(* IEC 61131-3 sources: plc-st-coding-agent/progress/evidence/f14_v3_parallel_20261112/jobs/custom_minimax-m27 (part 2) *)

(* ---- public-hard-06.candidate_01.st ---- *)
FUNCTION_BLOCK ProductionControl
VAR_INPUT
    Mode            : BOOL;
    ForwardButton   : BOOL;
    ReverseButton   : BOOL;
    SensorFeed      : BOOL;
    SensorWash      : BOOL;
    SensorWeight    : BOOL;
    SensorFiring    : BOOL;
    SensorOutput    : BOOL;
    washComplete    : BOOL;
    weightComplete  : BOOL;
    weight          : REAL;
    firingComplete  : BOOL;
END_VAR

VAR_OUTPUT
    MotorForward    : BOOL;
    MotorReverse    : BOOL;
    kick             : BOOL;
    CompletionLight  : BOOL;
    firingTemp       : REAL;
END_VAR

VAR
    State           : INT;
    prevSensorFeed  : BOOL;
    prevSensorWash  : BOOL;
    prevSensorWeight: BOOL;
    prevSensorFiring: BOOL;
    prevSensorOutput: BOOL;
END_VAR

TYPE ProductionState : INT (
    IDLE            := 0,
    MOVING_TO_WASH  := 1,
    AT_WASH         := 2,
    MOVING_TO_WEIGH := 3,
    AT_WEIGH        := 4,
    QUALITY_CHECK   := 5,
    KICKING         := 6,
    CALCULATING_TEMP:= 7,
    MOVING_TO_FIRING:= 8,
    AT_FIRING       := 9,
    MOVING_TO_OUTPUT:= 10,
    AT_OUTPUT       := 11
);
END_TYPE;

// Edge detection helpers
prevSensorFeed  := SensorFeed;
prevSensorWash  := SensorWash;
prevSensorWeight:= SensorWeight;
prevSensorFiring:= SensorFiring;
prevSensorOutput:= SensorOutput;

// Default outputs
MotorForward    := FALSE;
MotorReverse    := FALSE;
kick             := FALSE;
CompletionLight  := FALSE;
firingTemp       := 0.0;

IF Mode = FALSE THEN
    // Manual Mode
    IF ForwardButton AND NOT ReverseButton THEN
        MotorForward := TRUE;
        MotorReverse := FALSE;
    ELSIF ReverseButton AND NOT ForwardButton THEN
        MotorForward := FALSE;
        MotorReverse := TRUE;
    ELSE
        MotorForward := FALSE;
        MotorReverse := FALSE;
    END_IF;
    State := IDLE;
ELSE
    // Automatic Mode
    CASE State OF
        IDLE:
            IF SensorFeed AND NOT prevSensorFeed THEN
                State := MOVING_TO_WASH;
                MotorForward := TRUE;
            END_IF;

        MOVING_TO_WASH:
            IF SensorWash AND NOT prevSensorWash THEN
                State := AT_WASH;
                MotorForward := FALSE;
            END_IF;

        AT_WASH:
            IF washComplete THEN
                State := MOVING_TO_WEIGH;
                MotorForward := TRUE;
            END_IF;

        MOVING_TO_WEIGH:
            IF SensorWeight AND NOT prevSensorWeight THEN
                State := AT_WEIGH;
                MotorForward := FALSE;
            END_IF;

        AT_WEIGH:
            IF weightComplete THEN
                State := QUALITY_CHECK;
            END_IF;

        QUALITY_CHECK:
            IF weight < 100.0 OR weight > 200.0 THEN
                State := KICKING;
            ELSE
                State := CALCULATING_TEMP;
            END_IF;

        KICKING:
            kick := TRUE;
            State := IDLE;

        CALCULATING_TEMP:
            firingTemp := 500.0 + ((weight - 100.0) / 100.0) * 50.0;
            State := MOVING_TO_FIRING;
            MotorForward := TRUE;

        MOVING_TO_FIRING:
            IF SensorFiring AND NOT prevSensorFiring THEN
                State := AT_FIRING;
                MotorForward := FALSE;
            END_IF;

        AT_FIRING:
            IF firingComplete THEN
                State := MOVING_TO_OUTPUT;
                MotorForward := TRUE;
            END_IF;

        MOVING_TO_OUTPUT:
            IF SensorOutput AND NOT prevSensorOutput THEN
                State := AT_OUTPUT;
                MotorForward := FALSE;
            END_IF;

        AT_OUTPUT:
            CompletionLight := SensorOutput;
            IF NOT SensorOutput THEN
                State := IDLE;
                firingTemp := 0.0;
            END_IF;
    END_CASE;
END_IF;
END_FUNCTION_BLOCK

(* ---- public-hard-06.candidate_02.st ---- *)
FUNCTION_BLOCK ProductionControl
VAR_INPUT
    Mode            : BOOL;
    ForwardButton   : BOOL;
    ReverseButton   : BOOL;
    SensorFeed      : BOOL;
    SensorWash      : BOOL;
    SensorWeight    : BOOL;
    SensorFiring    : BOOL;
    SensorOutput    : BOOL;
    washComplete    : BOOL;
    weightComplete  : BOOL;
    weight          : REAL;
    firingComplete  : BOOL;
END_VAR

VAR_OUTPUT
    MotorForward    : BOOL;
    MotorReverse    : BOOL;
    kick             : BOOL;
    CompletionLight  : BOOL;
    firingTemp       : REAL;
END_VAR

VAR
    State           : INT;
    prevSensorFeed  : BOOL;
    prevSensorWash  : BOOL;
    prevSensorWeight: BOOL;
    prevSensorFiring: BOOL;
    prevSensorOutput: BOOL;
    prodState        : INT;
END_VAR

prodState := State;

kick := FALSE;
firingTemp := 0.0;

prevSensorFeed := SensorFeed;
prevSensorWash := SensorWash;
prevSensorWeight := SensorWeight;
prevSensorFiring := SensorFiring;
prevSensorOutput := SensorOutput;

IF Mode = FALSE THEN
    MotorForward := FALSE;
    MotorReverse := FALSE;
    kick := FALSE;
    CompletionLight := FALSE;
    IF ForwardButton AND NOT ReverseButton THEN
        MotorForward := TRUE;
    END_IF;
    IF ReverseButton AND NOT ForwardButton THEN
        MotorReverse := TRUE;
    END_IF;
    State := 0;
ELSE
    CompletionLight := FALSE;
    CASE State OF
        0:
            MotorForward := FALSE;
            MotorReverse := FALSE;
            kick := FALSE;
            IF SensorFeed AND NOT prevSensorFeed THEN
                State := 1;
            END_IF;

        1:
            MotorForward := TRUE;
            MotorReverse := FALSE;
            IF SensorWash AND NOT prevSensorWash THEN
                State := 2;
            END_IF;

        2:
            MotorForward := FALSE;
            MotorReverse := FALSE;
            IF washComplete THEN
                State := 3;
            END_IF;

        3:
            MotorForward := TRUE;
            MotorReverse := FALSE;
            IF SensorWeight AND NOT prevSensorWeight THEN
                State := 4;
            END_IF;

        4:
            MotorForward := FALSE;
            MotorReverse := FALSE;
            IF weightComplete THEN
                State := 5;
            END_IF;

        5:
            MotorForward := FALSE;
            MotorReverse := FALSE;
            IF weight < 100.0 OR weight > 200.0 THEN
                State := 6;
            ELSE
                State := 7;
            END_IF;

        6:
            kick := TRUE;
            MotorForward := FALSE;
            MotorReverse := FALSE;
            State := 0;

        7:
            kick := FALSE;
            firingTemp := 500.0 + ((weight - 100.0) / 100.0) * 50.0;
            State := 8;

        8:
            MotorForward := TRUE;
            MotorReverse := FALSE;
            kick := FALSE;
            IF SensorFiring AND NOT prevSensorFiring THEN
                State := 9;
            END_IF;

        9:
            MotorForward := FALSE;
            MotorReverse := FALSE;
            IF firingComplete THEN
                State := 10;
            END_IF;

        10:
            MotorForward := TRUE;
            MotorReverse := FALSE;
            IF SensorOutput AND NOT prevSensorOutput THEN
                State := 11;
            END_IF;

        11:
            MotorForward := FALSE;
            MotorReverse := FALSE;
            CompletionLight := TRUE;
            IF NOT SensorOutput THEN
                CompletionLight := FALSE;
                firingTemp := 0.0;
                State := 0;
            END_IF;
    END_CASE;
END_IF;
END_FUNCTION_BLOCK

(* ---- public-hard-06.raw_candidate_01.st ---- *)
FUNCTION_BLOCK ProductionControl
VAR_INPUT
    Mode            : BOOL;
    ForwardButton   : BOOL;
    ReverseButton   : BOOL;
    SensorFeed      : BOOL;
    SensorWash      : BOOL;
    SensorWeight    : BOOL;
    SensorFiring    : BOOL;
    SensorOutput    : BOOL;
    washComplete    : BOOL;
    weightComplete  : BOOL;
    weight          : REAL;
    firingComplete  : BOOL;
END_VAR

VAR_OUTPUT
    MotorForward    : BOOL;
    MotorReverse    : BOOL;
    kick             : BOOL;
    CompletionLight  : BOOL;
    firingTemp       : REAL;
END_VAR

VAR
    State           : INT;
    prevSensorFeed  : BOOL;
    prevSensorWash  : BOOL;
    prevSensorWeight: BOOL;
    prevSensorFiring: BOOL;
    prevSensorOutput: BOOL;
END_VAR

TYPE ProductionState : INT (
    IDLE            := 0,
    MOVING_TO_WASH  := 1,
    AT_WASH         := 2,
    MOVING_TO_WEIGH := 3,
    AT_WEIGH        := 4,
    QUALITY_CHECK   := 5,
    KICKING         := 6,
    CALCULATING_TEMP:= 7,
    MOVING_TO_FIRING:= 8,
    AT_FIRING       := 9,
    MOVING_TO_OUTPUT:= 10,
    AT_OUTPUT       := 11
);
END_TYPE

// Edge detection helpers
prevSensorFeed  := SensorFeed;
prevSensorWash  := SensorWash;
prevSensorWeight:= SensorWeight;
prevSensorFiring:= SensorFiring;
prevSensorOutput:= SensorOutput;

// Default outputs
MotorForward    := FALSE;
MotorReverse    := FALSE;
kick             := FALSE;
CompletionLight  := FALSE;
firingTemp       := 0.0;

IF Mode = FALSE THEN
    // Manual Mode
    IF ForwardButton AND NOT ReverseButton THEN
        MotorForward := TRUE;
        MotorReverse := FALSE;
    ELSIF ReverseButton AND NOT ForwardButton THEN
        MotorForward := FALSE;
        MotorReverse := TRUE;
    ELSE
        MotorForward := FALSE;
        MotorReverse := FALSE;
    END_IF;
    State := IDLE;
ELSE
    // Automatic Mode
    CASE State OF
        IDLE:
            IF SensorFeed AND NOT prevSensorFeed THEN
                State := MOVING_TO_WASH;
                MotorForward := TRUE;
            END_IF;

        MOVING_TO_WASH:
            IF SensorWash AND NOT prevSensorWash THEN
                State := AT_WASH;
                MotorForward := FALSE;
            END_IF;

        AT_WASH:
            IF washComplete THEN
                State := MOVING_TO_WEIGH;
                MotorForward := TRUE;
            END_IF;

        MOVING_TO_WEIGH:
            IF SensorWeight AND NOT prevSensorWeight THEN
                State := AT_WEIGH;
                MotorForward := FALSE;
            END_IF;

        AT_WEIGH:
            IF weightComplete THEN
                State := QUALITY_CHECK;
            END_IF;

        QUALITY_CHECK:
            IF weight < 100.0 OR weight > 200.0 THEN
                State := KICKING;
            ELSE
                State := CALCULATING_TEMP;
            END_IF;

        KICKING:
            kick := TRUE;
            State := IDLE;

        CALCULATING_TEMP:
            firingTemp := 500.0 + ((weight - 100.0) / 100.0) * 50.0;
            State := MOVING_TO_FIRING;
            MotorForward := TRUE;

        MOVING_TO_FIRING:
            IF SensorFiring AND NOT prevSensorFiring THEN
                State := AT_FIRING;
                MotorForward := FALSE;
            END_IF;

        AT_FIRING:
            IF firingComplete THEN
                State := MOVING_TO_OUTPUT;
                MotorForward := TRUE;
            END_IF;

        MOVING_TO_OUTPUT:
            IF SensorOutput AND NOT prevSensorOutput THEN
                State := AT_OUTPUT;
                MotorForward := FALSE;
            END_IF;

        AT_OUTPUT:
            CompletionLight := SensorOutput;
            IF NOT SensorOutput THEN
                State := IDLE;
                firingTemp := 0.0;
            END_IF;
    END_CASE;
END_IF;
END_FUNCTION_BLOCK

(* ---- public-hard-06.raw_candidate_02.st ---- *)
FUNCTION_BLOCK ProductionControl
VAR_INPUT
    Mode            : BOOL;
    ForwardButton   : BOOL;
    ReverseButton   : BOOL;
    SensorFeed      : BOOL;
    SensorWash      : BOOL;
    SensorWeight    : BOOL;
    SensorFiring    : BOOL;
    SensorOutput    : BOOL;
    washComplete    : BOOL;
    weightComplete  : BOOL;
    weight          : REAL;
    firingComplete  : BOOL;
END_VAR

VAR_OUTPUT
    MotorForward    : BOOL;
    MotorReverse    : BOOL;
    kick             : BOOL;
    CompletionLight  : BOOL;
    firingTemp       : REAL;
END_VAR

VAR
    State           : INT;
    prevSensorFeed  : BOOL;
    prevSensorWash  : BOOL;
    prevSensorWeight: BOOL;
    prevSensorFiring: BOOL;
    prevSensorOutput: BOOL;
    prodState        : INT;
END_VAR

prodState := State;

kick := FALSE;
firingTemp := 0.0;

prevSensorFeed := SensorFeed;
prevSensorWash := SensorWash;
prevSensorWeight := SensorWeight;
prevSensorFiring := SensorFiring;
prevSensorOutput := SensorOutput;

IF Mode = FALSE THEN
    MotorForward := FALSE;
    MotorReverse := FALSE;
    kick := FALSE;
    CompletionLight := FALSE;
    IF ForwardButton AND NOT ReverseButton THEN
        MotorForward := TRUE;
    END_IF;
    IF ReverseButton AND NOT ForwardButton THEN
        MotorReverse := TRUE;
    END_IF;
    State := 0;
ELSE
    CompletionLight := FALSE;
    CASE State OF
        0:
            MotorForward := FALSE;
            MotorReverse := FALSE;
            kick := FALSE;
            IF SensorFeed AND NOT prevSensorFeed THEN
                State := 1;
            END_IF;

        1:
            MotorForward := TRUE;
            MotorReverse := FALSE;
            IF SensorWash AND NOT prevSensorWash THEN
                State := 2;
            END_IF;

        2:
            MotorForward := FALSE;
            MotorReverse := FALSE;
            IF washComplete THEN
                State := 3;
            END_IF;

        3:
            MotorForward := TRUE;
            MotorReverse := FALSE;
            IF SensorWeight AND NOT prevSensorWeight THEN
                State := 4;
            END_IF;

        4:
            MotorForward := FALSE;
            MotorReverse := FALSE;
            IF weightComplete THEN
                State := 5;
            END_IF;

        5:
            MotorForward := FALSE;
            MotorReverse := FALSE;
            IF weight < 100.0 OR weight > 200.0 THEN
                State := 6;
            ELSE
                State := 7;
            END_IF;

        6:
            kick := TRUE;
            MotorForward := FALSE;
            MotorReverse := FALSE;
            State := 0;

        7:
            kick := FALSE;
            firingTemp := 500.0 + ((weight - 100.0) / 100.0) * 50.0;
            State := 8;

        8:
            MotorForward := TRUE;
            MotorReverse := FALSE;
            kick := FALSE;
            IF SensorFiring AND NOT prevSensorFiring THEN
                State := 9;
            END_IF;

        9:
            MotorForward := FALSE;
            MotorReverse := FALSE;
            IF firingComplete THEN
                State := 10;
            END_IF;

        10:
            MotorForward := TRUE;
            MotorReverse := FALSE;
            IF SensorOutput AND NOT prevSensorOutput THEN
                State := 11;
            END_IF;

        11:
            MotorForward := FALSE;
            MotorReverse := FALSE;
            CompletionLight := TRUE;
            IF NOT SensorOutput THEN
                CompletionLight := FALSE;
                firingTemp := 0.0;
                State := 0;
            END_IF;
    END_CASE;
END_IF;
END_FUNCTION_BLOCK

(* ---- public-medium-01.candidate_01.st ---- *)
FUNCTION_BLOCK FB_MultiPumpControl
VAR_INPUT
    mode  : BOOL;    // FALSE: Manual, TRUE: Automatic
    start : BOOL;    // Start button
    stop  : BOOL;    // Stop button
END_VAR

VAR_IN_OUT
    pumpGroup : ARRAY[1..5] OF ST_Pump;
END_VAR

VAR
    lastStart : BOOL := FALSE;
    lastStop  : BOOL := FALSE;
    edgeStart : BOOL;
    edgeStop  : BOOL;
    i         : INT;
    j         : INT;
    tempPri   : INT;
    tempSel   : BOOL;
    tempCmd   : BOOL;
    sorted    : ARRAY[1..5] OF ST_Pump;
END_VAR

// Edge detection for rising edges
edgeStart := start AND NOT lastStart;
edgeStop  := stop  AND NOT lastStop;
lastStart := start;
lastStop  := stop;

// Stop all pumps when stop button is pressed
IF edgeStop THEN
    FOR i := 1 TO 5 DO
        pumpGroup[i].RunComd := FALSE;
    END_FOR;
END_IF;

// Start selected pumps when start button is pressed
IF edgeStart THEN
    IF mode = FALSE THEN
        // Manual mode: run pumps where selection = TRUE
        FOR i := 1 TO 5 DO
            pumpGroup[i].RunComd := pumpGroup[i].selection;
        END_FOR;
    ELSE
        // Automatic mode: three pumps in use, two on standby
        // Sort pumps by priority (descending) using bubble sort
        sorted := pumpGroup;
        FOR i := 1 TO 4 DO
            FOR j := 1 TO 5 - i DO
                IF sorted[j].priority < sorted[j + 1].priority THEN
                    tempPri := sorted[j].priority;
                    tempSel := sorted[j].selection;
                    tempCmd := sorted[j].RunComd;
                    sorted[j].priority   := sorted[j + 1].priority;
                    sorted[j].selection  := sorted[j + 1].selection;
                    sorted[j].RunComd    := sorted[j + 1].RunComd;
                    sorted[j + 1].priority := tempPri;
                    sorted[j + 1].selection := tempSel;
                    sorted[j + 1].RunComd   := tempCmd;
                END_IF;
            END_FOR;
        END_FOR;
        // Top 3 highest priority pumps run
        sorted[1].RunComd := TRUE;
        sorted[2].RunComd := TRUE;
        sorted[3].RunComd := TRUE;
        sorted[4].RunComd := FALSE;
        sorted[5].RunComd := FALSE;
        // Copy RunComd back to original array (preserving original order)
        FOR i := 1 TO 5 DO
            pumpGroup[i].RunComd := sorted[i].RunComd;
        END_FOR;
    END_IF;
END_IF;

END_FUNCTION_BLOCK

(* ---- public-medium-01.candidate_02.st ---- *)
TYPE ST_Pump : STRUCT
    priority : INT;
    selection : BOOL;
    runCmd   : BOOL;
END_STRUCT;
END_TYPE;

FUNCTION_BLOCK FB_MultiPumpControl
VAR_INPUT
    mode  : BOOL;
    start : BOOL;
    stop  : BOOL;
END_VAR

VAR_IN_OUT
    pumpGroup : ARRAY[1..5] OF ST_Pump;
END_VAR

VAR
    lastStart : BOOL := FALSE;
    lastStop  : BOOL := FALSE;
    edgeStart : BOOL;
    edgeStop  : BOOL;
    i         : INT;
    j         : INT;
    tempPump  : ST_Pump;
    pumpSorted : ARRAY[1..5] OF ST_Pump;
END_VAR

edgeStart := start AND NOT lastStart;
edgeStop  := stop  AND NOT lastStop;
lastStart := start;
lastStop  := stop;

IF edgeStop THEN
    FOR i := 1 TO 5 DO
        pumpGroup[i].runCmd := FALSE;
    END_FOR;
END_IF;

IF edgeStart THEN
    IF mode = FALSE THEN
        FOR i := 1 TO 5 DO
            pumpGroup[i].runCmd := pumpGroup[i].selection;
        END_FOR;
    ELSE
        pumpSorted := pumpGroup;
        FOR i := 1 TO 4 DO
            FOR j := 1 TO 5 - i DO
                IF pumpSorted[j].priority < pumpSorted[j + 1].priority THEN
                    tempPump := pumpSorted[j];
                    pumpSorted[j] := pumpSorted[j + 1];
                    pumpSorted[j + 1] := tempPump;
                END_IF;
            END_FOR;
        END_FOR;
        pumpSorted[1].runCmd := TRUE;
        pumpSorted[2].runCmd := TRUE;
        pumpSorted[3].runCmd := TRUE;
        pumpSorted[4].runCmd := FALSE;
        pumpSorted[5].runCmd := FALSE;
        pumpGroup := pumpSorted;
    END_IF;
END_IF;

END_FUNCTION_BLOCK

(* ---- public-medium-01.raw_candidate_01.st ---- *)
FUNCTION_BLOCK FB_MultiPumpControl
VAR_INPUT
    mode  : BOOL;    // FALSE: Manual, TRUE: Automatic
    start : BOOL;    // Start button
    stop  : BOOL;    // Stop button
END_VAR

VAR_IN_OUT
    pumpGroup : ARRAY[1..5] OF ST_Pump;
END_VAR

VAR
    lastStart : BOOL := FALSE;
    lastStop  : BOOL := FALSE;
    edgeStart : BOOL;
    edgeStop  : BOOL;
    i         : INT;
    j         : INT;
    tempPri   : INT;
    tempSel   : BOOL;
    tempCmd   : BOOL;
    sorted    : ARRAY[1..5] OF ST_Pump;
END_VAR

// Edge detection for rising edges
edgeStart := start AND NOT lastStart;
edgeStop  := stop  AND NOT lastStop;
lastStart := start;
lastStop  := stop;

// Stop all pumps when stop button is pressed
IF edgeStop THEN
    FOR i := 1 TO 5 DO
        pumpGroup[i].RunComd := FALSE;
    END_FOR;
END_IF

// Start selected pumps when start button is pressed
IF edgeStart THEN
    IF mode = FALSE THEN
        // Manual mode: run pumps where selection = TRUE
        FOR i := 1 TO 5 DO
            pumpGroup[i].RunComd := pumpGroup[i].selection;
        END_FOR;
    ELSE
        // Automatic mode: three pumps in use, two on standby
        // Sort pumps by priority (descending) using bubble sort
        sorted := pumpGroup;
        FOR i := 1 TO 4 DO
            FOR j := 1 TO 5 - i DO
                IF sorted[j].priority < sorted[j + 1].priority THEN
                    tempPri := sorted[j].priority;
                    tempSel := sorted[j].selection;
                    tempCmd := sorted[j].RunComd;
                    sorted[j].priority   := sorted[j + 1].priority;
                    sorted[j].selection  := sorted[j + 1].selection;
                    sorted[j].RunComd    := sorted[j + 1].RunComd;
                    sorted[j + 1].priority := tempPri;
                    sorted[j + 1].selection := tempSel;
                    sorted[j + 1].RunComd   := tempCmd;
                END_IF
            END_FOR
        END_FOR
        // Top 3 highest priority pumps run
        sorted[1].RunComd := TRUE;
        sorted[2].RunComd := TRUE;
        sorted[3].RunComd := TRUE;
        sorted[4].RunComd := FALSE;
        sorted[5].RunComd := FALSE;
        // Copy RunComd back to original array (preserving original order)
        FOR i := 1 TO 5 DO
            pumpGroup[i].RunComd := sorted[i].RunComd;
        END_FOR;
    END_IF
END_IF

END_FUNCTION_BLOCK

(* ---- public-medium-01.raw_candidate_02.st ---- *)
TYPE ST_Pump : STRUCT
    priority : INT;
    selection : BOOL;
    runCmd   : BOOL;
END_STRUCT
END_TYPE

FUNCTION_BLOCK FB_MultiPumpControl
VAR_INPUT
    mode  : BOOL;
    start : BOOL;
    stop  : BOOL;
END_VAR

VAR_IN_OUT
    pumpGroup : ARRAY[1..5] OF ST_Pump;
END_VAR

VAR
    lastStart : BOOL := FALSE;
    lastStop  : BOOL := FALSE;
    edgeStart : BOOL;
    edgeStop  : BOOL;
    i         : INT;
    j         : INT;
    tempPump  : ST_Pump;
    pumpSorted : ARRAY[1..5] OF ST_Pump;
END_VAR

edgeStart := start AND NOT lastStart;
edgeStop  := stop  AND NOT lastStop;
lastStart := start;
lastStop  := stop;

IF edgeStop THEN
    FOR i := 1 TO 5 DO
        pumpGroup[i].runCmd := FALSE;
    END_FOR;
END_IF;

IF edgeStart THEN
    IF mode = FALSE THEN
        FOR i := 1 TO 5 DO
            pumpGroup[i].runCmd := pumpGroup[i].selection;
        END_FOR;
    ELSE
        pumpSorted := pumpGroup;
        FOR i := 1 TO 4 DO
            FOR j := 1 TO 5 - i DO
                IF pumpSorted[j].priority < pumpSorted[j + 1].priority THEN
                    tempPump := pumpSorted[j];
                    pumpSorted[j] := pumpSorted[j + 1];
                    pumpSorted[j + 1] := tempPump;
                END_IF;
            END_FOR;
        END_FOR;
        pumpSorted[1].runCmd := TRUE;
        pumpSorted[2].runCmd := TRUE;
        pumpSorted[3].runCmd := TRUE;
        pumpSorted[4].runCmd := FALSE;
        pumpSorted[5].runCmd := FALSE;
        pumpGroup := pumpSorted;
    END_IF;
END_IF;

END_FUNCTION_BLOCK

(* ---- public-medium-02.candidate_01.st ---- *)
FUNCTION_BLOCK FB_AnalogBatchProcessing
VAR_INPUT
    count : DINT;
END_VAR

VAR_IN_OUT
    analogValues : ARRAY[*] OF INT;
    channels : ARRAY[*] OF ST_AnalogChannel;
END_VAR

VAR
    i : DINT;
    idx : DINT;
    rawValue : INT;
    rawMin : INT;
    rawMax : INT;
    loLIM : REAL;
    hiLIM : REAL;
END_VAR

loLIM := 0.0;
hiLIM := 0.0;

FOR i := 0 TO count - 1 DO
    idx := LOWER_BOUND(analogValues, 1) + i;
    rawValue := analogValues[idx];

    channels[idx].retVal := 16#0000;

    IF channels[idx].enable THEN
        loLIM := channels[idx].loLIM;
        hiLIM := channels[idx].hiLIM;

        CASE channels[idx].measuringMode OF
            0: // Non-temperature linear scaling
                IF hiLIM > loLIM THEN
                    IF channels[idx].bipolar THEN
                        rawMin := -27648;
                        rawMax := 27648;
                    ELSE
                        rawMin := 0;
                        rawMax := 27648;
                    END_IF;

                    channels[idx].outputValue := TO_REAL(rawValue - rawMin) / TO_REAL(rawMax - rawMin) * (hiLIM - loLIM) + loLIM;
                ELSE
                    channels[idx].retVal := 16#8002;
                END_IF;

            1: // Standard temperature: outputValue = raw / 10
                channels[idx].outputValue := TO_REAL(rawValue) / 10.0;

            2: // Climatic temperature: outputValue = raw / 100
                channels[idx].outputValue := TO_REAL(rawValue) / 100.0;

            ELSE
                channels[idx].retVal := 16#8001;
        END_CASE;
    END_IF;
END_FOR;
END_FUNCTION_BLOCK

(* ---- public-medium-02.candidate_02.st ---- *)
TYPE ST_AnalogChannel :
STRUCT
    enable : BOOL;
    hiLIM : REAL;
    loLIM : REAL;
    bipolar : BOOL;
    measuringMode : INT;
    retVal : WORD;
    outputValue : REAL;
END_STRUCT;
END_TYPE;

FUNCTION_BLOCK FB_AnalogBatchProcessing
VAR_INPUT
    count : DINT;
END_VAR

VAR_IN_OUT
    analogValues : ARRAY[*] OF INT;
    channels : ARRAY[*] OF ST_AnalogChannel;
END_VAR

VAR
    i : DINT;
    idx : DINT;
    rawValue : INT;
    rawMin : INT;
    rawMax : INT;
    chLoLIM : REAL;
    chHiLIM : REAL;
    ch : REFERENCE TO ST_AnalogChannel;
END_VAR

FOR i := 0 TO count - 1 DO
    idx := LOWER_BOUND(analogValues, 1) + i;
    rawValue := analogValues[idx];
    ch REF= channels[idx];
    ch.retVal := 16#0000;

    IF ch.enable THEN
        chLoLIM := ch.loLIM;
        chHiLIM := ch.hiLIM;

        CASE ch.measuringMode OF
            0:
                IF chHiLIM > chLoLIM THEN
                    IF ch.bipolar THEN
                        rawMin := -27648;
                        rawMax := 27648;
                    ELSE
                        rawMin := 0;
                        rawMax := 27648;
                    END_IF;
                    ch.outputValue := INT_TO_REAL(rawValue - rawMin) / INT_TO_REAL(rawMax - rawMin) * (chHiLIM - chLoLIM) + chLoLIM;
                ELSE
                    ch.retVal := 16#8002;
                END_IF;

            1:
                ch.outputValue := INT_TO_REAL(rawValue) / 10.0;

            2:
                ch.outputValue := INT_TO_REAL(rawValue) / 100.0;

            ELSE
                ch.retVal := 16#8001;
        END_CASE;
    END_IF;
END_FOR;
END_FUNCTION_BLOCK

(* ---- public-medium-02.raw_candidate_01.st ---- *)
FUNCTION_BLOCK FB_AnalogBatchProcessing
VAR_INPUT
    count : DINT;
END_VAR

VAR_IN_OUT
    analogValues : ARRAY[*] OF INT;
    channels : ARRAY[*] OF ST_AnalogChannel;
END_VAR

VAR
    i : DINT;
    idx : DINT;
    rawValue : INT;
    rawMin : INT;
    rawMax : INT;
    loLIM : REAL;
    hiLIM : REAL;
END_VAR

loLIM := 0.0;
hiLIM := 0.0;

FOR i := 0 TO count - 1 DO
    idx := LOWER_BOUND(analogValues, 1) + i;
    rawValue := analogValues[idx];

    channels[idx].retVal := 16#0000;

    IF channels[idx].enable THEN
        loLIM := channels[idx].loLIM;
        hiLIM := channels[idx].hiLIM;

        CASE channels[idx].measuringMode OF
            0: // Non-temperature linear scaling
                IF hiLIM > loLIM THEN
                    IF channels[idx].bipolar THEN
                        rawMin := -27648;
                        rawMax := 27648;
                    ELSE
                        rawMin := 0;
                        rawMax := 27648;
                    END_IF;

                    channels[idx].outputValue := TO_REAL(rawValue - rawMin) / TO_REAL(rawMax - rawMin) * (hiLIM - loLIM) + loLIM;
                ELSE
                    channels[idx].retVal := 16#8002;
                END_IF;

            1: // Standard temperature: outputValue = raw / 10
                channels[idx].outputValue := TO_REAL(rawValue) / 10.0;

            2: // Climatic temperature: outputValue = raw / 100
                channels[idx].outputValue := TO_REAL(rawValue) / 100.0;

            ELSE
                channels[idx].retVal := 16#8001;
        END_CASE;
    END_IF;
END_FOR;
END_FUNCTION_BLOCK

(* ---- public-medium-02.raw_candidate_02.st ---- *)
TYPE ST_AnalogChannel :
STRUCT
    enable : BOOL;
    hiLIM : REAL;
    loLIM : REAL;
    bipolar : BOOL;
    measuringMode : INT;
    retVal : WORD;
    outputValue : REAL;
END_STRUCT
END_TYPE

FUNCTION_BLOCK FB_AnalogBatchProcessing
VAR_INPUT
    count : DINT;
END_VAR

VAR_IN_OUT
    analogValues : ARRAY[*] OF INT;
    channels : ARRAY[*] OF ST_AnalogChannel;
END_VAR

VAR
    i : DINT;
    idx : DINT;
    rawValue : INT;
    rawMin : INT;
    rawMax : INT;
    chLoLIM : REAL;
    chHiLIM : REAL;
    ch : REFERENCE TO ST_AnalogChannel;
END_VAR

FOR i := 0 TO count - 1 DO
    idx := LOWER_BOUND(analogValues, 1) + i;
    rawValue := analogValues[idx];
    ch REF= channels[idx];
    ch.retVal := 16#0000;

    IF ch.enable THEN
        chLoLIM := ch.loLIM;
        chHiLIM := ch.hiLIM;

        CASE ch.measuringMode OF
            0:
                IF chHiLIM > chLoLIM THEN
                    IF ch.bipolar THEN
                        rawMin := -27648;
                        rawMax := 27648;
                    ELSE
                        rawMin := 0;
                        rawMax := 27648;
                    END_IF;
                    ch.outputValue := INT_TO_REAL(rawValue - rawMin) / INT_TO_REAL(rawMax - rawMin) * (chHiLIM - chLoLIM) + chLoLIM;
                ELSE
                    ch.retVal := 16#8002;
                END_IF;

            1:
                ch.outputValue := INT_TO_REAL(rawValue) / 10.0;

            2:
                ch.outputValue := INT_TO_REAL(rawValue) / 100.0;

            ELSE
                ch.retVal := 16#8001;
        END_CASE;
    END_IF;
END_FOR;
END_FUNCTION_BLOCK

(* ---- public-medium-03.candidate_01.st ---- *)
FUNCTION_BLOCK FB_MovingAverage
VAR_INPUT
    cyclicExecution : BOOL;
    trigger : BOOL;
    value : LREAL;
    windowSize : INT;
    reset : BOOL;
END_VAR

VAR_OUTPUT
    average : LREAL;
    windowSizeReached : BOOL;
    error : BOOL;
    status : WORD;
END_VAR

VAR
    dataBuffer : ARRAY[1..100] OF LREAL;
    sum : LREAL;
    count : INT;
    writeIndex : INT;
    lastTrigger : BOOL;
    lastReset : BOOL;
    initValid : BOOL;
END_VAR

// Reset handling
IF reset AND NOT lastReset THEN
    sum := 0.0;
    count := 0;
    writeIndex := 0;
    average := 0.0;
    windowSizeReached := FALSE;
    error := FALSE;
    status := 16#0000;
    initValid := FALSE;
END_IF;
lastReset := reset;

// Validate window size on first execution or when reset was just released
IF NOT initValid THEN
    IF windowSize < 1 OR windowSize > 100 THEN
        error := TRUE;
        status := 16#8200;
        RETURN;
    ELSE
        error := FALSE;
        status := 16#0000;
        initValid := TRUE;
    END_IF;
END_IF;

// Check for cyclic execution mode
IF cyclicExecution THEN
    // Validate window size on each cycle
    IF windowSize < 1 OR windowSize > 100 THEN
        error := TRUE;
        status := 16#8200;
        RETURN;
    ELSE
        error := FALSE;
        status := 16#0000;
    END_IF;

    // Process new value
    IF count >= windowSize THEN
        sum := sum - dataBuffer[writeIndex + 1];
    ELSE
        count := count + 1;
    END_IF;

    writeIndex := (writeIndex MOD windowSize) + 1;
    dataBuffer[writeIndex] := value;
    sum := sum + value;

    IF count >= windowSize THEN
        windowSizeReached := TRUE;
    ELSE
        windowSizeReached := FALSE;
    END_IF;

    average := sum / INT_TO_LREAL(count);
    lastTrigger := FALSE;
    RETURN;
END_IF;

// Check for rising edge on trigger
IF trigger AND NOT lastTrigger THEN
    // Validate window size
    IF windowSize < 1 OR windowSize > 100 THEN
        error := TRUE;
        status := 16#8200;
        lastTrigger := trigger;
        RETURN;
    ELSE
        error := FALSE;
        status := 16#0000;
    END_IF;

    // Process new value
    IF count >= windowSize THEN
        sum := sum - dataBuffer[writeIndex + 1];
    ELSE
        count := count + 1;
    END_IF;

    writeIndex := (writeIndex MOD windowSize) + 1;
    dataBuffer[writeIndex] := value;
    sum := sum + value;

    IF count >= windowSize THEN
        windowSizeReached := TRUE;
    ELSE
        windowSizeReached := FALSE;
    END_IF;

    average := sum / INT_TO_LREAL(count);
END_IF;

lastTrigger := trigger;
END_FUNCTION_BLOCK

(* ---- public-medium-03.candidate_02.st ---- *)
FUNCTION_BLOCK FB_MovingAverage
VAR_INPUT
    cyclicExecution : BOOL;
    trigger : BOOL;
    value : LREAL;
    windowSize : INT;
    reset : BOOL;
END_VAR

VAR_OUTPUT
    average : LREAL;
    windowSizeReached : BOOL;
    error : BOOL;
    status : WORD;
END_VAR

VAR
    dataBuffer : ARRAY[1..100] OF LREAL;
    sum : LREAL;
    count : INT;
    writeIndex : INT;
    lastTrigger : BOOL;
    lastReset : BOOL;
    initValid : BOOL;
END_VAR

IF reset AND NOT lastReset THEN
    sum := 0.0;
    count := 0;
    writeIndex := 0;
    average := 0.0;
    windowSizeReached := FALSE;
    error := FALSE;
    status := 16#0000;
    initValid := FALSE;
END_IF;
lastReset := reset;

IF NOT initValid THEN
    IF windowSize < 1 OR windowSize > 100 THEN
        error := TRUE;
        status := 16#8200;
        RETURN;
    ELSE
        error := FALSE;
        status := 16#0000;
        initValid := TRUE;
    END_IF;
END_IF;

IF cyclicExecution THEN
    IF windowSize < 1 OR windowSize > 100 THEN
        error := TRUE;
        status := 16#8200;
        RETURN;
    ELSE
        error := FALSE;
        status := 16#0000;
    END_IF;

    IF count >= windowSize THEN
        sum := sum - dataBuffer[((writeIndex) MOD windowSize) + 1];
    ELSE
        count := count + 1;
    END_IF;

    writeIndex := writeIndex + 1;
    IF writeIndex > windowSize THEN
        writeIndex := 1;
    END_IF;

    dataBuffer[writeIndex] := value;
    sum := sum + value;

    IF count >= windowSize THEN
        windowSizeReached := TRUE;
        average := sum / INT_TO_LREAL(windowSize);
    ELSE
        windowSizeReached := FALSE;
        average := sum / INT_TO_LREAL(count);
    END_IF;
    lastTrigger := FALSE;
    RETURN;
END_IF;

IF trigger AND NOT lastTrigger THEN
    IF windowSize < 1 OR windowSize > 100 THEN
        error := TRUE;
        status := 16#8200;
        lastTrigger := trigger;
        RETURN;
    ELSE
        error := FALSE;
        status := 16#0000;
    END_IF;

    IF count >= windowSize THEN
        sum := sum - dataBuffer[((writeIndex) MOD windowSize) + 1];
    ELSE
        count := count + 1;
    END_IF;

    writeIndex := writeIndex + 1;
    IF writeIndex > windowSize THEN
        writeIndex := 1;
    END_IF;

    dataBuffer[writeIndex] := value;
    sum := sum + value;

    IF count >= windowSize THEN
        windowSizeReached := TRUE;
        average := sum / INT_TO_LREAL(windowSize);
    ELSE
        windowSizeReached := FALSE;
        average := sum / INT_TO_LREAL(count);
    END_IF;
END_IF;

lastTrigger := trigger;
END_FUNCTION_BLOCK

(* ---- public-medium-03.raw_candidate_01.st ---- *)
FUNCTION_BLOCK FB_MovingAverage
VAR_INPUT
    cyclicExecution : BOOL;
    trigger : BOOL;
    value : LREAL;
    windowSize : INT;
    reset : BOOL;
END_VAR

VAR_OUTPUT
    average : LREAL;
    windowSizeReached : BOOL;
    error : BOOL;
    status : WORD;
END_VAR

VAR
    dataBuffer : ARRAY[1..100] OF LREAL;
    sum : LREAL;
    count : INT;
    writeIndex : INT;
    lastTrigger : BOOL;
    lastReset : BOOL;
    initValid : BOOL;
END_VAR

// Reset handling
IF reset AND NOT lastReset THEN
    sum := 0.0;
    count := 0;
    writeIndex := 0;
    average := 0.0;
    windowSizeReached := FALSE;
    error := FALSE;
    status := 16#0000;
    initValid := FALSE;
END_IF;
lastReset := reset;

// Validate window size on first execution or when reset was just released
IF NOT initValid THEN
    IF windowSize < 1 OR windowSize > 100 THEN
        error := TRUE;
        status := 16#8200;
        RETURN;
    ELSE
        error := FALSE;
        status := 16#0000;
        initValid := TRUE;
    END_IF;
END_IF;

// Check for cyclic execution mode
IF cyclicExecution THEN
    // Validate window size on each cycle
    IF windowSize < 1 OR windowSize > 100 THEN
        error := TRUE;
        status := 16#8200;
        RETURN;
    ELSE
        error := FALSE;
        status := 16#0000;
    END_IF;

    // Process new value
    IF count >= windowSize THEN
        sum := sum - dataBuffer[writeIndex + 1];
    ELSE
        count := count + 1;
    END_IF;

    writeIndex := (writeIndex MOD windowSize) + 1;
    dataBuffer[writeIndex] := value;
    sum := sum + value;

    IF count >= windowSize THEN
        windowSizeReached := TRUE;
    ELSE
        windowSizeReached := FALSE;
    END_IF;

    average := sum / INT_TO_LREAL(count);
    lastTrigger := FALSE;
    RETURN;
END_IF;

// Check for rising edge on trigger
IF trigger AND NOT lastTrigger THEN
    // Validate window size
    IF windowSize < 1 OR windowSize > 100 THEN
        error := TRUE;
        status := 16#8200;
        lastTrigger := trigger;
        RETURN;
    ELSE
        error := FALSE;
        status := 16#0000;
    END_IF;

    // Process new value
    IF count >= windowSize THEN
        sum := sum - dataBuffer[writeIndex + 1];
    ELSE
        count := count + 1;
    END_IF;

    writeIndex := (writeIndex MOD windowSize) + 1;
    dataBuffer[writeIndex] := value;
    sum := sum + value;

    IF count >= windowSize THEN
        windowSizeReached := TRUE;
    ELSE
        windowSizeReached := FALSE;
    END_IF;

    average := sum / INT_TO_LREAL(count);
END_IF;

lastTrigger := trigger;
END_FUNCTION_BLOCK

(* ---- public-medium-03.raw_candidate_02.st ---- *)
FUNCTION_BLOCK FB_MovingAverage
VAR_INPUT
    cyclicExecution : BOOL;
    trigger : BOOL;
    value : LREAL;
    windowSize : INT;
    reset : BOOL;
END_VAR

VAR_OUTPUT
    average : LREAL;
    windowSizeReached : BOOL;
    error : BOOL;
    status : WORD;
END_VAR

VAR
    dataBuffer : ARRAY[1..100] OF LREAL;
    sum : LREAL;
    count : INT;
    writeIndex : INT;
    lastTrigger : BOOL;
    lastReset : BOOL;
    initValid : BOOL;
END_VAR

IF reset AND NOT lastReset THEN
    sum := 0.0;
    count := 0;
    writeIndex := 0;
    average := 0.0;
    windowSizeReached := FALSE;
    error := FALSE;
    status := 16#0000;
    initValid := FALSE;
END_IF;
lastReset := reset;

IF NOT initValid THEN
    IF windowSize < 1 OR windowSize > 100 THEN
        error := TRUE;
        status := 16#8200;
        RETURN;
    ELSE
        error := FALSE;
        status := 16#0000;
        initValid := TRUE;
    END_IF;
END_IF;

IF cyclicExecution THEN
    IF windowSize < 1 OR windowSize > 100 THEN
        error := TRUE;
        status := 16#8200;
        RETURN;
    ELSE
        error := FALSE;
        status := 16#0000;
    END_IF;

    IF count >= windowSize THEN
        sum := sum - dataBuffer[((writeIndex) MOD windowSize) + 1];
    ELSE
        count := count + 1;
    END_IF;

    writeIndex := writeIndex + 1;
    IF writeIndex > windowSize THEN
        writeIndex := 1;
    END_IF;

    dataBuffer[writeIndex] := value;
    sum := sum + value;

    IF count >= windowSize THEN
        windowSizeReached := TRUE;
        average := sum / INT_TO_LREAL(windowSize);
    ELSE
        windowSizeReached := FALSE;
        average := sum / INT_TO_LREAL(count);
    END_IF;
    lastTrigger := FALSE;
    RETURN;
END_IF;

IF trigger AND NOT lastTrigger THEN
    IF windowSize < 1 OR windowSize > 100 THEN
        error := TRUE;
        status := 16#8200;
        lastTrigger := trigger;
        RETURN;
    ELSE
        error := FALSE;
        status := 16#0000;
    END_IF;

    IF count >= windowSize THEN
        sum := sum - dataBuffer[((writeIndex) MOD windowSize) + 1];
    ELSE
        count := count + 1;
    END_IF;

    writeIndex := writeIndex + 1;
    IF writeIndex > windowSize THEN
        writeIndex := 1;
    END_IF;

    dataBuffer[writeIndex] := value;
    sum := sum + value;

    IF count >= windowSize THEN
        windowSizeReached := TRUE;
        average := sum / INT_TO_LREAL(windowSize);
    ELSE
        windowSizeReached := FALSE;
        average := sum / INT_TO_LREAL(count);
    END_IF;
END_IF;

lastTrigger := trigger;
END_FUNCTION_BLOCK

(* ---- public-medium-04.candidate_01.st ---- *)
FUNCTION_BLOCK FB_TemperatureControl
VAR_INPUT
    TemperatureSensorInput : REAL;
    SetTemperature : REAL;
END_VAR
VAR_OUTPUT
    CurrentTemperature : REAL;
    SetTempDisplay : REAL;
    HeaterStatus : BOOL;
    OverheatProtection : BOOL;
    HeaterOutput : BOOL;
END_VAR
VAR
    OverheatTimer : TON;
    LockoutTimer : TON;
    OverheatTriggered : BOOL := FALSE;
    LockoutActive : BOOL := FALSE;
END_VAR

(* Constants *)
OverheatTimer.PT := T#5S;
LockoutTimer.PT := T#3S;

(* Sensor fault check: temperature out of valid range *)
IF TemperatureSensorInput < 0.0 OR TemperatureSensorInput > 100.0 THEN
    HeaterOutput := FALSE;
    OverheatTimer(IN := FALSE);
    LockoutTimer(IN := FALSE);
    LockoutActive := FALSE;
    OverheatTriggered := FALSE;
ELSE
    (* Normal temperature control *)

    (* Start overheat timer when heater is commanded ON *)
    OverheatTimer(IN := TRUE);

    (* Check if overheat timer exceeded 5s → trigger protection *)
    IF OverheatTimer.Q AND NOT OverheatTriggered THEN
        OverheatTriggered := TRUE;
        LockoutActive := TRUE;
        LockoutTimer(IN := TRUE);
    END_IF;

    (* If protection triggered, force heater OFF and wait lockout *)
    IF OverheatTriggered THEN
        HeaterOutput := FALSE;

        (* After lockout expires, clear protection *)
        IF LockoutTimer.Q THEN
            LockoutActive := FALSE;
            OverheatTriggered := FALSE;
            LockoutTimer(IN := FALSE);
            OverheatTimer(IN := FALSE);
        END_IF;
    ELSE
        (* Normal operation: compare temperature vs setpoint *)
        IF TemperatureSensorInput < SetTemperature THEN
            HeaterOutput := TRUE;
        ELSE
            HeaterOutput := FALSE;
        END_IF;
    END_IF;

    (* Reset overheat timer when heater is OFF (but not in protection) *)
    IF NOT HeaterOutput AND NOT OverheatTriggered THEN
        OverheatTimer(IN := FALSE);
    END_IF;
END_IF;

(* Update display outputs *)
CurrentTemperature := TemperatureSensorInput;
SetTempDisplay := SetTemperature;
HeaterStatus := HeaterOutput;
OverheatProtection := OverheatTriggered;

END_FUNCTION_BLOCK

(* ---- public-medium-04.candidate_02.st ---- *)
FUNCTION_BLOCK FB_TemperatureControl
VAR_INPUT
    TemperatureSensorInput : REAL;
    SetTemperature : REAL;
END_VAR
VAR_OUTPUT
    CurrentTemperature : REAL;
    SetTempDisplay : REAL;
    HeaterStatus : BOOL;
    OverheatProtection : BOOL;
    HeaterOutput : BOOL;
END_VAR
VAR
    OverheatTimer : TON;
    LockoutTimer : TON;
    OverheatTriggered : BOOL := FALSE;
END_VAR

OverheatTimer.PT := T#5S;
LockoutTimer.PT := T#3S;

(* Sensor fault check: temperature out of valid range *)
IF TemperatureSensorInput < 0.0 OR TemperatureSensorInput > 100.0 THEN
    HeaterOutput := FALSE;
    OverheatTimer(IN := FALSE);
    LockoutTimer(IN := FALSE);
    OverheatTimer(IN := FALSE, PT := T#5S);
    OverheatTriggered := FALSE;
ELSE
    (* Normal temperature control *)
    IF NOT OverheatTriggered THEN
        (* Normal heating decision *)
        IF TemperatureSensorInput < SetTemperature THEN
            HeaterOutput := TRUE;
        ELSE
            HeaterOutput := FALSE;
        END_IF;
    ELSE
        (* Overheat protection active - heater forced off *)
        HeaterOutput := FALSE;
    END_IF;

    (* Overheat timer: accumulate time only when heater is ON and not in protection *)
    IF NOT OverheatTriggered AND HeaterOutput THEN
        OverheatTimer(IN := TRUE);
    ELSE
        OverheatTimer(IN := FALSE);
    END_IF;

    (* Check overheat threshold *)
    IF OverheatTimer.Q AND NOT OverheatTriggered THEN
        OverheatTriggered := TRUE;
    END_IF;

    (* Lockout timer management *)
    IF OverheatTriggered THEN
        LockoutTimer(IN := TRUE);
        IF LockoutTimer.Q THEN
            OverheatTriggered := FALSE;
            LockoutTimer(IN := FALSE);
            OverheatTimer(IN := FALSE, PT := T#5S);
        END_IF;
    ELSE
        LockoutTimer(IN := FALSE);
    END_IF;
END_IF;

(* Update display outputs *)
CurrentTemperature := TemperatureSensorInput;
SetTempDisplay := SetTemperature;
HeaterStatus := HeaterOutput;
OverheatProtection := OverheatTriggered;

END_FUNCTION_BLOCK

(* ---- public-medium-04.raw_candidate_01.st ---- *)
FUNCTION_BLOCK FB_TemperatureControl
VAR_INPUT
    TemperatureSensorInput : REAL;
    SetTemperature : REAL;
END_VAR
VAR_OUTPUT
    CurrentTemperature : REAL;
    SetTempDisplay : REAL;
    HeaterStatus : BOOL;
    OverheatProtection : BOOL;
    HeaterOutput : BOOL;
END_VAR
VAR
    OverheatTimer : TON;
    LockoutTimer : TON;
    OverheatTriggered : BOOL := FALSE;
    LockoutActive : BOOL := FALSE;
END_VAR

(* Constants *)
OverheatTimer.PT := T#5S;
LockoutTimer.PT := T#3S;

(* Sensor fault check: temperature out of valid range *)
IF TemperatureSensorInput < 0.0 OR TemperatureSensorInput > 100.0 THEN
    HeaterOutput := FALSE;
    OverheatTimer(IN := FALSE);
    LockoutTimer(IN := FALSE);
    LockoutActive := FALSE;
    OverheatTriggered := FALSE;
ELSE
    (* Normal temperature control *)

    (* Start overheat timer when heater is commanded ON *)
    OverheatTimer(IN := TRUE);

    (* Check if overheat timer exceeded 5s → trigger protection *)
    IF OverheatTimer.Q AND NOT OverheatTriggered THEN
        OverheatTriggered := TRUE;
        LockoutActive := TRUE;
        LockoutTimer(IN := TRUE);
    END_IF

    (* If protection triggered, force heater OFF and wait lockout *)
    IF OverheatTriggered THEN
        HeaterOutput := FALSE;

        (* After lockout expires, clear protection *)
        IF LockoutTimer.Q THEN
            LockoutActive := FALSE;
            OverheatTriggered := FALSE;
            LockoutTimer(IN := FALSE);
            OverheatTimer(IN := FALSE);
        END_IF
    ELSE
        (* Normal operation: compare temperature vs setpoint *)
        IF TemperatureSensorInput < SetTemperature THEN
            HeaterOutput := TRUE;
        ELSE
            HeaterOutput := FALSE;
        END_IF
    END_IF

    (* Reset overheat timer when heater is OFF (but not in protection) *)
    IF NOT HeaterOutput AND NOT OverheatTriggered THEN
        OverheatTimer(IN := FALSE);
    END_IF
END_IF

(* Update display outputs *)
CurrentTemperature := TemperatureSensorInput;
SetTempDisplay := SetTemperature;
HeaterStatus := HeaterOutput;
OverheatProtection := OverheatTriggered;

END_FUNCTION_BLOCK

(* ---- public-medium-04.raw_candidate_02.st ---- *)
FUNCTION_BLOCK FB_TemperatureControl
VAR_INPUT
    TemperatureSensorInput : REAL;
    SetTemperature : REAL;
END_VAR
VAR_OUTPUT
    CurrentTemperature : REAL;
    SetTempDisplay : REAL;
    HeaterStatus : BOOL;
    OverheatProtection : BOOL;
    HeaterOutput : BOOL;
END_VAR
VAR
    OverheatTimer : TON;
    LockoutTimer : TON;
    OverheatTriggered : BOOL := FALSE;
END_VAR

OverheatTimer.PT := T#5S;
LockoutTimer.PT := T#3S;

(* Sensor fault check: temperature out of valid range *)
IF TemperatureSensorInput < 0.0 OR TemperatureSensorInput > 100.0 THEN
    HeaterOutput := FALSE;
    OverheatTimer(IN := FALSE);
    LockoutTimer(IN := FALSE);
    OverheatTimer(IN := FALSE, PT := T#5S);
    OverheatTriggered := FALSE;
ELSE
    (* Normal temperature control *)
    IF NOT OverheatTriggered THEN
        (* Normal heating decision *)
        IF TemperatureSensorInput < SetTemperature THEN
            HeaterOutput := TRUE;
        ELSE
            HeaterOutput := FALSE;
        END_IF;
    ELSE
        (* Overheat protection active - heater forced off *)
        HeaterOutput := FALSE;
    END_IF;

    (* Overheat timer: accumulate time only when heater is ON and not in protection *)
    IF NOT OverheatTriggered AND HeaterOutput THEN
        OverheatTimer(IN := TRUE);
    ELSE
        OverheatTimer(IN := FALSE);
    END_IF;

    (* Check overheat threshold *)
    IF OverheatTimer.Q AND NOT OverheatTriggered THEN
        OverheatTriggered := TRUE;
    END_IF;

    (* Lockout timer management *)
    IF OverheatTriggered THEN
        LockoutTimer(IN := TRUE);
        IF LockoutTimer.Q THEN
            OverheatTriggered := FALSE;
            LockoutTimer(IN := FALSE);
            OverheatTimer(IN := FALSE, PT := T#5S);
        END_IF;
    ELSE
        LockoutTimer(IN := FALSE);
    END_IF;
END_IF;

(* Update display outputs *)
CurrentTemperature := TemperatureSensorInput;
SetTempDisplay := SetTemperature;
HeaterStatus := HeaterOutput;
OverheatProtection := OverheatTriggered;

END_FUNCTION_BLOCK

(* ---- public-medium-05.candidate_01.st ---- *)
TYPE ProdState :
(
    WAIT_A      : UINT := 0,
    STAGE_A     : UINT := 1,
    MOVING_AB   : UINT := 2,
    STAGE_B     : UINT := 3,
    MOVING_BC   : UINT := 4,
    STAGE_C     : UINT := 5,
    COMPLETE    : UINT := 6
);
END_TYPE;

FUNCTION_BLOCK ProductionLineControl
VAR
    State : ProdState := WAIT_A;
    NextState : ProdState;
END_VAR
VAR_OUTPUT
    MotorForward    : BOOL;
    MotorReverse    : BOOL;
    CompletionLight : BOOL;
END_VAR

NextState := State;

IF Mode = FALSE THEN
    // Manual Mode
    MotorForward  := ForwardButton AND NOT ReverseButton;
    MotorReverse  := ReverseButton AND NOT ForwardButton;
    NextState     := WAIT_A;
ELSE
    // Automatic Mode
    MotorForward  := FALSE;
    MotorReverse  := FALSE;

    IF State = WAIT_A THEN
        IF SensorA THEN
            NextState := STAGE_A;
        END_IF;
    ELSIF State = STAGE_A THEN
        IF SensorA AND ButtonA THEN
            NextState := MOVING_AB;
        END_IF;
    ELSIF State = MOVING_AB THEN
        MotorForward := TRUE;
        IF SensorB THEN
            NextState := STAGE_B;
        END_IF;
    ELSIF State = STAGE_B THEN
        IF SensorB AND ButtonB THEN
            NextState := MOVING_BC;
        END_IF;
    ELSIF State = MOVING_BC THEN
        MotorForward := TRUE;
        IF SensorC THEN
            NextState := STAGE_C;
        END_IF;
    ELSIF State = STAGE_C THEN
        IF SensorC AND ButtonC THEN
            NextState := COMPLETE;
        END_IF;
    ELSIF State = COMPLETE THEN
        IF NOT SensorC THEN
            NextState := WAIT_A;
        END_IF;
    END_IF;
END_IF;

State := NextState;

CompletionLight := (State = COMPLETE) AND SensorC;

END_FUNCTION_BLOCK

(* ---- public-medium-05.candidate_02.st ---- *)
TYPE ProdState : (WAIT_A, STAGE_A, MOVING_AB, STAGE_B, MOVING_BC, STAGE_C, COMPLETE);
END_TYPE;

FUNCTION_BLOCK ProductionLineControl
VAR
    State : ProdState := WAIT_A;
    NextState : ProdState;
END_VAR
VAR_OUTPUT
    MotorForward    : BOOL;
    MotorReverse    : BOOL;
    CompletionLight : BOOL;
END_VAR

NextState := State;

IF Mode = FALSE THEN
    MotorForward  := ForwardButton AND NOT ReverseButton;
    MotorReverse  := ReverseButton AND NOT ForwardButton;
    NextState     := WAIT_A;
ELSE
    MotorForward  := FALSE;
    MotorReverse  := FALSE;
    CASE State OF
        WAIT_A:
            IF SensorA THEN
                NextState := STAGE_A;
            END_IF;
        STAGE_A:
            IF SensorA AND ButtonA THEN
                NextState := MOVING_AB;
            END_IF;
        MOVING_AB:
            MotorForward := TRUE;
            IF SensorB THEN
                NextState := STAGE_B;
            END_IF;
        STAGE_B:
            IF SensorB AND ButtonB THEN
                NextState := MOVING_BC;
            END_IF;
        MOVING_BC:
            MotorForward := TRUE;
            IF SensorC THEN
                NextState := STAGE_C;
            END_IF;
        STAGE_C:
            IF SensorC AND ButtonC THEN
                NextState := COMPLETE;
            END_IF;
        COMPLETE:
            IF NOT SensorC THEN
                NextState := WAIT_A;
            END_IF;
    END_CASE;
END_IF;

State := NextState;

CompletionLight := (State = COMPLETE) AND SensorC;

END_FUNCTION_BLOCK

(* ---- public-medium-05.raw_candidate_01.st ---- *)
TYPE ProdState :
(
    WAIT_A      : UINT := 0,
    STAGE_A     : UINT := 1,
    MOVING_AB   : UINT := 2,
    STAGE_B     : UINT := 3,
    MOVING_BC   : UINT := 4,
    STAGE_C     : UINT := 5,
    COMPLETE    : UINT := 6
);
END_TYPE

FUNCTION_BLOCK ProductionLineControl
VAR
    State : ProdState := WAIT_A;
    NextState : ProdState;
END_VAR
VAR_OUTPUT
    MotorForward    : BOOL;
    MotorReverse    : BOOL;
    CompletionLight : BOOL;
END_VAR

NextState := State;

IF Mode = FALSE THEN
    // Manual Mode
    MotorForward  := ForwardButton AND NOT ReverseButton;
    MotorReverse  := ReverseButton AND NOT ForwardButton;
    NextState     := WAIT_A;
ELSE
    // Automatic Mode
    MotorForward  := FALSE;
    MotorReverse  := FALSE;

    IF State = WAIT_A THEN
        IF SensorA THEN
            NextState := STAGE_A;
        END_IF
    ELSIF State = STAGE_A THEN
        IF SensorA AND ButtonA THEN
            NextState := MOVING_AB;
        END_IF
    ELSIF State = MOVING_AB THEN
        MotorForward := TRUE;
        IF SensorB THEN
            NextState := STAGE_B;
        END_IF
    ELSIF State = STAGE_B THEN
        IF SensorB AND ButtonB THEN
            NextState := MOVING_BC;
        END_IF
    ELSIF State = MOVING_BC THEN
        MotorForward := TRUE;
        IF SensorC THEN
            NextState := STAGE_C;
        END_IF
    ELSIF State = STAGE_C THEN
        IF SensorC AND ButtonC THEN
            NextState := COMPLETE;
        END_IF
    ELSIF State = COMPLETE THEN
        IF NOT SensorC THEN
            NextState := WAIT_A;
        END_IF
    END_IF;
END_IF;

State := NextState;

CompletionLight := (State = COMPLETE) AND SensorC;

END_FUNCTION_BLOCK

(* ---- public-medium-05.raw_candidate_02.st ---- *)
TYPE ProdState : (WAIT_A, STAGE_A, MOVING_AB, STAGE_B, MOVING_BC, STAGE_C, COMPLETE);
END_TYPE

FUNCTION_BLOCK ProductionLineControl
VAR
    State : ProdState := WAIT_A;
    NextState : ProdState;
END_VAR
VAR_OUTPUT
    MotorForward    : BOOL;
    MotorReverse    : BOOL;
    CompletionLight : BOOL;
END_VAR

NextState := State;

IF Mode = FALSE THEN
    MotorForward  := ForwardButton AND NOT ReverseButton;
    MotorReverse  := ReverseButton AND NOT ForwardButton;
    NextState     := WAIT_A;
ELSE
    MotorForward  := FALSE;
    MotorReverse  := FALSE;
    CASE State OF
        WAIT_A:
            IF SensorA THEN
                NextState := STAGE_A;
            END_IF;
        STAGE_A:
            IF SensorA AND ButtonA THEN
                NextState := MOVING_AB;
            END_IF;
        MOVING_AB:
            MotorForward := TRUE;
            IF SensorB THEN
                NextState := STAGE_B;
            END_IF;
        STAGE_B:
            IF SensorB AND ButtonB THEN
                NextState := MOVING_BC;
            END_IF;
        MOVING_BC:
            MotorForward := TRUE;
            IF SensorC THEN
                NextState := STAGE_C;
            END_IF;
        STAGE_C:
            IF SensorC AND ButtonC THEN
                NextState := COMPLETE;
            END_IF;
        COMPLETE:
            IF NOT SensorC THEN
                NextState := WAIT_A;
            END_IF;
    END_CASE;
END_IF;

State := NextState;

CompletionLight := (State = COMPLETE) AND SensorC;

END_FUNCTION_BLOCK

(* ---- public-medium-06.candidate_01.st ---- *)
FUNCTION_BLOCK SlabThicknessMonitor
VAR_INPUT
    THICKNESS_FAULT        : BOOL;
    THICKNESS_SIGNAL_VALID : BOOL;
    CUTTING_RUN            : BOOL;
    FaultTimestamp         : DINT;
    CycleTime              : TIME;
END_VAR

VAR_OUTPUT
    THICKNESS_ALARM          : BOOL;
    Slab_Fault_Counter       : UINT;
    Slab_Runtime_Accumulator : LTIME;
    Slab_Fault_History       : ARRAY[0..4] OF DINT;
END_VAR

VAR
    AlarmHoldTimer    : TON;
    PreviousFaultValid : BOOL;
    FirstScan          : BOOL;
    i                  : INT;
END_VAR

// Power-up initialization
IF FirstScan THEN
    FirstScan := FALSE;
    Slab_Fault_Counter := 0;
    Slab_Runtime_Accumulator := LTIME#0;
    FOR i := 0 TO 4 DO
        Slab_Fault_History[i] := 0;
    END_FOR;
END_IF;

// Signal validity: clears alarm/hold state and blocks all processing
IF NOT THICKNESS_SIGNAL_VALID THEN
    THICKNESS_ALARM := FALSE;
    AlarmHoldTimer(IN := FALSE);
    PreviousFaultValid := FALSE;
ELSE
    // Rising edge detection of valid fault signal
    IF THICKNESS_FAULT AND NOT PreviousFaultValid THEN
        Slab_Fault_Counter := Slab_Fault_Counter + 1;
        FOR i := 4 TO 1 BY -1 DO
            Slab_Fault_History[i] := Slab_Fault_History[i-1];
        END_FOR;
        Slab_Fault_History[0] := FaultTimestamp;
    END_IF;
    PreviousFaultValid := THICKNESS_FAULT;

    // Runtime accumulation
    IF CUTTING_RUN AND NOT THICKNESS_FAULT THEN
        Slab_Runtime_Accumulator := Slab_Runtime_Accumulator + CycleTime;
    END_IF;

    // Alarm activation and 500 ms hold logic
    IF THICKNESS_FAULT THEN
        THICKNESS_ALARM := TRUE;
        AlarmHoldTimer(IN := FALSE);
    ELSIF THICKNESS_ALARM AND NOT AlarmHoldTimer.Q THEN
        AlarmHoldTimer(IN := TRUE, PT := T#500ms);
    ELSIF NOT AlarmHoldTimer.Q THEN
        THICKNESS_ALARM := FALSE;
    END_IF;
END_IF;
END_FUNCTION_BLOCK

(* ---- public-medium-06.candidate_02.st ---- *)
FUNCTION_BLOCK SlabThicknessMonitor
VAR_INPUT
    THICKNESS_FAULT        : BOOL;
    THICKNESS_SIGNAL_VALID : BOOL;
    CUTTING_RUN            : BOOL;
    FaultTimestamp         : DINT;
    CycleTime              : TIME;
END_VAR

VAR_OUTPUT
    THICKNESS_ALARM          : BOOL;
    Slab_Fault_Counter       : UINT;
    Slab_Runtime_Accumulator : LTIME;
    Slab_Fault_History       : ARRAY[0..4] OF DINT;
END_VAR

VAR
    AlarmHoldTimer     : TON;
    PreviousFaultValid : BOOL;
    FirstScan          : BOOL;
    idx                : INT;
END_VAR

IF FirstScan THEN
    FirstScan := FALSE;
    Slab_Fault_Counter := 0;
    Slab_Runtime_Accumulator := LTIME#0ms;
    FOR idx := 0 TO 4 DO
        Slab_Fault_History[idx] := 0;
    END_FOR;
END_IF;

IF NOT THICKNESS_SIGNAL_VALID THEN
    THICKNESS_ALARM := FALSE;
    AlarmHoldTimer(IN := FALSE);
    PreviousFaultValid := FALSE;
ELSE
    IF THICKNESS_FAULT AND NOT PreviousFaultValid THEN
        Slab_Fault_Counter := Slab_Fault_Counter + 1;
        FOR idx := 4 TO 1 BY -1 DO
            Slab_Fault_History[idx] := Slab_Fault_History[idx-1];
        END_FOR;
        Slab_Fault_History[0] := FaultTimestamp;
    END_IF;
    PreviousFaultValid := THICKNESS_FAULT;

    IF CUTTING_RUN AND NOT THICKNESS_FAULT THEN
        Slab_Runtime_Accumulator := Slab_Runtime_Accumulator + TO_LTIME(CycleTime);
    END_IF;

    IF THICKNESS_FAULT THEN
        THICKNESS_ALARM := TRUE;
        AlarmHoldTimer(IN := FALSE);
    ELSIF THICKNESS_ALARM AND NOT AlarmHoldTimer.Q THEN
        AlarmHoldTimer(IN := TRUE, PT := T#500ms);
    ELSIF NOT AlarmHoldTimer.Q THEN
        THICKNESS_ALARM := FALSE;
    END_IF;
END_IF;
END_FUNCTION_BLOCK

(* ---- public-medium-06.raw_candidate_01.st ---- *)
FUNCTION_BLOCK SlabThicknessMonitor
VAR_INPUT
    THICKNESS_FAULT        : BOOL;
    THICKNESS_SIGNAL_VALID : BOOL;
    CUTTING_RUN            : BOOL;
    FaultTimestamp         : DINT;
    CycleTime              : TIME;
END_VAR

VAR_OUTPUT
    THICKNESS_ALARM          : BOOL;
    Slab_Fault_Counter       : UINT;
    Slab_Runtime_Accumulator : LTIME;
    Slab_Fault_History       : ARRAY[0..4] OF DINT;
END_VAR

VAR
    AlarmHoldTimer    : TON;
    PreviousFaultValid : BOOL;
    FirstScan          : BOOL;
    i                  : INT;
END_VAR

// Power-up initialization
IF FirstScan THEN
    FirstScan := FALSE;
    Slab_Fault_Counter := 0;
    Slab_Runtime_Accumulator := LTIME#0;
    FOR i := 0 TO 4 DO
        Slab_Fault_History[i] := 0;
    END_FOR;
END_IF;

// Signal validity: clears alarm/hold state and blocks all processing
IF NOT THICKNESS_SIGNAL_VALID THEN
    THICKNESS_ALARM := FALSE;
    AlarmHoldTimer(IN := FALSE);
    PreviousFaultValid := FALSE;
ELSE
    // Rising edge detection of valid fault signal
    IF THICKNESS_FAULT AND NOT PreviousFaultValid THEN
        Slab_Fault_Counter := Slab_Fault_Counter + 1;
        FOR i := 4 TO 1 BY -1 DO
            Slab_Fault_History[i] := Slab_Fault_History[i-1];
        END_FOR;
        Slab_Fault_History[0] := FaultTimestamp;
    END_IF;
    PreviousFaultValid := THICKNESS_FAULT;

    // Runtime accumulation
    IF CUTTING_RUN AND NOT THICKNESS_FAULT THEN
        Slab_Runtime_Accumulator := Slab_Runtime_Accumulator + CycleTime;
    END_IF;

    // Alarm activation and 500 ms hold logic
    IF THICKNESS_FAULT THEN
        THICKNESS_ALARM := TRUE;
        AlarmHoldTimer(IN := FALSE);
    ELSIF THICKNESS_ALARM AND NOT AlarmHoldTimer.Q THEN
        AlarmHoldTimer(IN := TRUE, PT := T#500ms);
    ELSIF NOT AlarmHoldTimer.Q THEN
        THICKNESS_ALARM := FALSE;
    END_IF;
END_IF;
END_FUNCTION_BLOCK

(* ---- public-medium-06.raw_candidate_02.st ---- *)
FUNCTION_BLOCK SlabThicknessMonitor
VAR_INPUT
    THICKNESS_FAULT        : BOOL;
    THICKNESS_SIGNAL_VALID : BOOL;
    CUTTING_RUN            : BOOL;
    FaultTimestamp         : DINT;
    CycleTime              : TIME;
END_VAR

VAR_OUTPUT
    THICKNESS_ALARM          : BOOL;
    Slab_Fault_Counter       : UINT;
    Slab_Runtime_Accumulator : LTIME;
    Slab_Fault_History       : ARRAY[0..4] OF DINT;
END_VAR

VAR
    AlarmHoldTimer     : TON;
    PreviousFaultValid : BOOL;
    FirstScan          : BOOL;
    idx                : INT;
END_VAR

IF FirstScan THEN
    FirstScan := FALSE;
    Slab_Fault_Counter := 0;
    Slab_Runtime_Accumulator := LTIME#0ms;
    FOR idx := 0 TO 4 DO
        Slab_Fault_History[idx] := 0;
    END_FOR;
END_IF;

IF NOT THICKNESS_SIGNAL_VALID THEN
    THICKNESS_ALARM := FALSE;
    AlarmHoldTimer(IN := FALSE);
    PreviousFaultValid := FALSE;
ELSE
    IF THICKNESS_FAULT AND NOT PreviousFaultValid THEN
        Slab_Fault_Counter := Slab_Fault_Counter + 1;
        FOR idx := 4 TO 1 BY -1 DO
            Slab_Fault_History[idx] := Slab_Fault_History[idx-1];
        END_FOR;
        Slab_Fault_History[0] := FaultTimestamp;
    END_IF;
    PreviousFaultValid := THICKNESS_FAULT;

    IF CUTTING_RUN AND NOT THICKNESS_FAULT THEN
        Slab_Runtime_Accumulator := Slab_Runtime_Accumulator + TO_LTIME(CycleTime);
    END_IF;

    IF THICKNESS_FAULT THEN
        THICKNESS_ALARM := TRUE;
        AlarmHoldTimer(IN := FALSE);
    ELSIF THICKNESS_ALARM AND NOT AlarmHoldTimer.Q THEN
        AlarmHoldTimer(IN := TRUE, PT := T#500ms);
    ELSIF NOT AlarmHoldTimer.Q THEN
        THICKNESS_ALARM := FALSE;
    END_IF;
END_IF;
END_FUNCTION_BLOCK

(* ---- public-medium-07.candidate_01.st ---- *)
FUNCTION_BLOCK HVAC_Control
VAR_INPUT
    OCCUPANCY_DETECTED    : BOOL;
    ENERGY_SAVING_MODE    : BOOL;
    HVAC_MODE_SELECTOR    : INT;
END_VAR

VAR_OUTPUT
    SUPPLY_FAN_RUN        : BOOL := FALSE;
    TEMP_SETPOINT_ADJUST  : INT := 0;
END_VAR

VAR
    fanDelayTimer : TON;
    fanConditionsMet : BOOL;
    rawAdjustment : INT;
END_VAR

(* Fan delay logic: 30s on, instant off *)
fanConditionsMet := OCCUPANCY_DETECTED AND (HVAC_MODE_SELECTOR <> 3);

fanDelayTimer(
    IN  := fanConditionsMet,
    PT  := T#30S
);

IF fanDelayTimer.Q THEN
    SUPPLY_FAN_RUN := TRUE;
ELSE
    SUPPLY_FAN_RUN := FALSE;
END_IF;

(* Temperature setpoint calculation *)
rawAdjustment := 0;

CASE HVAC_MODE_SELECTOR OF
    0: (* Auto mode *)
        IF OCCUPANCY_DETECTED THEN
            rawAdjustment := 0;
        ELSE
            IF ENERGY_SAVING_MODE THEN
                rawAdjustment := 3;
            ELSE
                rawAdjustment := 2;
            END_IF;
        END_IF;

    1: (* Comfort mode *)
        IF OCCUPANCY_DETECTED THEN
            rawAdjustment := 0;
        ELSE
            rawAdjustment := 1;
        END_IF;

    2: (* Economy mode *)
        IF OCCUPANCY_DETECTED THEN
            rawAdjustment := 0;
        ELSE
            rawAdjustment := 4;
        END_IF;

    3: (* Night mode *)
        rawAdjustment := 4;

ELSE
    rawAdjustment := 0;
END_CASE;

(* Clamp to ±4°C *)
IF rawAdjustment > 4 THEN
    TEMP_SETPOINT_ADJUST := 4;
ELSIF rawAdjustment < -4 THEN
    TEMP_SETPOINT_ADJUST := -4;
ELSE
    TEMP_SETPOINT_ADJUST := rawAdjustment;
END_IF;

END_FUNCTION_BLOCK

(* ---- public-medium-07.raw_candidate_01.st ---- *)
FUNCTION_BLOCK HVAC_Control
VAR_INPUT
    OCCUPANCY_DETECTED    : BOOL;
    ENERGY_SAVING_MODE    : BOOL;
    HVAC_MODE_SELECTOR    : INT;
END_VAR

VAR_OUTPUT
    SUPPLY_FAN_RUN        : BOOL := FALSE;
    TEMP_SETPOINT_ADJUST  : INT := 0;
END_VAR

VAR
    fanDelayTimer : TON;
    fanConditionsMet : BOOL;
    rawAdjustment : INT;
END_VAR

(* Fan delay logic: 30s on, instant off *)
fanConditionsMet := OCCUPANCY_DETECTED AND (HVAC_MODE_SELECTOR <> 3);

fanDelayTimer(
    IN  := fanConditionsMet,
    PT  := T#30S
);

IF fanDelayTimer.Q THEN
    SUPPLY_FAN_RUN := TRUE;
ELSE
    SUPPLY_FAN_RUN := FALSE;
END_IF;

(* Temperature setpoint calculation *)
rawAdjustment := 0;

CASE HVAC_MODE_SELECTOR OF
    0: (* Auto mode *)
        IF OCCUPANCY_DETECTED THEN
            rawAdjustment := 0;
        ELSE
            IF ENERGY_SAVING_MODE THEN
                rawAdjustment := 3;
            ELSE
                rawAdjustment := 2;
            END_IF;
        END_IF;

    1: (* Comfort mode *)
        IF OCCUPANCY_DETECTED THEN
            rawAdjustment := 0;
        ELSE
            rawAdjustment := 1;
        END_IF;

    2: (* Economy mode *)
        IF OCCUPANCY_DETECTED THEN
            rawAdjustment := 0;
        ELSE
            rawAdjustment := 4;
        END_IF;

    3: (* Night mode *)
        rawAdjustment := 4;

ELSE
    rawAdjustment := 0;
END_CASE;

(* Clamp to ±4°C *)
IF rawAdjustment > 4 THEN
    TEMP_SETPOINT_ADJUST := 4;
ELSIF rawAdjustment < -4 THEN
    TEMP_SETPOINT_ADJUST := -4;
ELSE
    TEMP_SETPOINT_ADJUST := rawAdjustment;
END_IF;

END_FUNCTION_BLOCK

(* ---- public-medium-08.candidate_01.st ---- *)
FUNCTION_BLOCK FB_ParseIPv4
VAR_INPUT
    ipText : STRING(254);
END_VAR
VAR_OUTPUT
    ipValue : UDINT;
END_VAR
VAR
    i : UINT;
    dot1 : UINT;
    dot2 : UINT;
    dot3 : UINT;
    len : UINT;
    seg1 : STRING(4);
    seg2 : STRING(4);
    seg3 : STRING(4);
    seg4 : STRING(4);
    seg1Len : UINT;
    seg2Len : UINT;
    seg3Len : UINT;
    seg4Len : UINT;
    val1 : UDINT;
    val2 : UDINT;
    val3 : UDINT;
    val4 : UDINT;
    result : UDINT;
    valid : BOOL;
    ch : CHAR;
END_VAR

result := 0;
valid := TRUE;

len := LEN(ipText);

IF len = 0 OR len > 254 THEN
    valid := FALSE;
END_IF;

IF valid THEN
    dot1 := FIND(ipText, '.');
    IF dot1 <= 1 OR dot1 >= 254 THEN
        valid := FALSE;
    END_IF;
END_IF;

IF valid THEN
    dot2 := FIND(MID(ipText, 254 - dot1, dot1 + 1), '.');
    IF dot2 > 0 THEN
        dot2 := dot2 + dot1;
    END_IF;
END_IF;

IF valid THEN
    dot3 := 0;
    IF dot2 > 0 AND dot2 < 254 THEN
        dot3 := FIND(MID(ipText, 254 - dot2, dot2 + 1), '.');
        IF dot3 > 0 THEN
            dot3 := dot3 + dot2;
        END_IF;
    END_IF;
END_IF;

IF valid THEN
    IF dot1 = 0 OR dot2 = 0 OR dot3 = 0 THEN
        valid := FALSE;
    END_IF;
END_IF;

IF valid THEN
    seg1Len := dot1 - 1;
    seg2Len := dot2 - dot1 - 1;
    seg3Len := dot3 - dot2 - 1;
    seg4Len := len - dot3;

    IF seg1Len < 1 OR seg1Len > 3 OR seg2Len < 1 OR seg2Len > 3 OR
       seg3Len < 1 OR seg3Len > 3 OR seg4Len < 1 OR seg4Len > 3 THEN
        valid := FALSE;
    END_IF;
END_IF;

IF valid THEN
    seg1 := LEFT(ipText, seg1Len);
    seg2 := MID(ipText, seg2Len, dot1 + 1);
    seg3 := MID(ipText, seg3Len, dot2 + 1);
    seg4 := RIGHT(ipText, seg4Len);

    valid := (seg1Len = LEN(seg1)) AND (seg2Len = LEN(seg2)) AND
             (seg3Len = LEN(seg3)) AND (seg4Len = LEN(seg4));
END_IF;

IF valid THEN
    valid := FALSE;
    val1 := STRING_TO_UDINT(seg1);
    val2 := STRING_TO_UDINT(seg2);
    val3 := STRING_TO_UDINT(seg3);
    val4 := STRING_TO_UDINT(seg4);

    FOR i := 1 TO seg1Len DO
        ch := MID(seg1, 1, i);
        IF (ch < '0') OR (ch > '9') THEN
            valid := TRUE;
        END_IF;
    END_FOR;

    IF NOT valid THEN
        FOR i := 1 TO seg2Len DO
            ch := MID(seg2, 1, i);
            IF (ch < '0') OR (ch > '9') THEN
                valid := TRUE;
            END_IF;
        END_FOR;
    END_IF;

    IF NOT valid THEN
        FOR i := 1 TO seg3Len DO
            ch := MID(seg3, 1, i);
            IF (ch < '0') OR (ch > '9') THEN
                valid := TRUE;
            END_IF;
        END_FOR;
    END_IF;

    IF NOT valid THEN
        FOR i := 1 TO seg4Len DO
            ch := MID(seg4, 1, i);
            IF (ch < '0') OR (ch > '9') THEN
                valid := TRUE;
            END_IF;
        END_FOR;
    END_IF;

    IF valid THEN
        valid := FALSE;
    END_IF;
END_IF;

IF valid THEN
    IF val1 <= 255 AND val2 <= 255 AND val3 <= 255 AND val4 <= 255 THEN
        result := (val1 * 16#1000000) OR (val2 * 16#10000) OR (val3 * 16#100) OR val4;
    END_IF;
END_IF;

ipValue := result;
END_FUNCTION_BLOCK

(* ---- public-medium-08.candidate_02.st ---- *)
FUNCTION_BLOCK FB_ParseIPv4
VAR_INPUT
    ipText : STRING(254);
END_VAR
VAR_OUTPUT
    ipValue : UDINT;
END_VAR
VAR
    i : UINT;
    dot1 : UINT;
    dot2 : UINT;
    dot3 : UINT;
    len : UINT;
    seg1 : STRING(4);
    seg2 : STRING(4);
    seg3 : STRING(4);
    seg4 : STRING(4);
    seg1Len : UINT;
    seg2Len : UINT;
    seg3Len : UINT;
    seg4Len : UINT;
    val1 : UDINT;
    val2 : UDINT;
    val3 : UDINT;
    val4 : UDINT;
    result : UDINT;
    valid : BOOL;
    ch : STRING(1);
END_VAR

result := 0;
valid := TRUE;

len := TO_UINT(LEN(ipText));

IF len = 0 OR len > 15 THEN
    valid := FALSE;
END_IF;

IF valid THEN
    dot1 := TO_UINT(FIND(ipText, '.'));
    IF dot1 <= 1 OR dot1 >= 254 THEN
        valid := FALSE;
    END_IF;
END_IF;

IF valid THEN
    dot2 := TO_UINT(FIND(MID(ipText, TO_INT(len - dot1), TO_INT(dot1 + 1)), '.'));
    IF dot2 > 0 THEN
        dot2 := dot2 + dot1;
    END_IF;
END_IF;

IF valid THEN
    dot3 := 0;
    IF dot2 > 0 AND dot2 < 254 THEN
        dot3 := TO_UINT(FIND(MID(ipText, TO_INT(len - dot2), TO_INT(dot2 + 1)), '.'));
        IF dot3 > 0 THEN
            dot3 := dot3 + dot2;
        END_IF;
    END_IF;
END_IF;

IF valid THEN
    IF dot1 = 0 OR dot2 = 0 OR dot3 = 0 THEN
        valid := FALSE;
    END_IF;
END_IF;

IF valid THEN
    seg1Len := dot1 - 1;
    seg2Len := dot2 - dot1 - 1;
    seg3Len := dot3 - dot2 - 1;
    seg4Len := len - dot3;

    IF seg1Len < 1 OR seg1Len > 3 OR seg2Len < 1 OR seg2Len > 3 OR seg3Len < 1 OR seg3Len > 3 OR seg4Len < 1 OR seg4Len > 3 THEN
        valid := FALSE;
    END_IF;
END_IF;

IF valid THEN
    seg1 := LEFT(ipText, TO_INT(seg1Len));
    seg2 := MID(ipText, TO_INT(seg2Len), TO_INT(dot1 + 1));
    seg3 := MID(ipText, TO_INT(seg3Len), TO_INT(dot2 + 1));
    seg4 := RIGHT(ipText, TO_INT(seg4Len));

    IF TO_UINT(LEN(seg1)) <> seg1Len OR TO_UINT(LEN(seg2)) <> seg2Len OR
       TO_UINT(LEN(seg3)) <> seg3Len OR TO_UINT(LEN(seg4)) <> seg4Len THEN
        valid := FALSE;
    END_IF;
END_IF;

IF valid THEN
    val1 := STRING_TO_UDINT(seg1);
    val2 := STRING_TO_UDINT(seg2);
    val3 := STRING_TO_UDINT(seg3);
    val4 := STRING_TO_UDINT(seg4);

    FOR i := 1 TO TO_INT(seg1Len) DO
        ch := MID(seg1, 1, TO_INT(i));
        IF ch < '0' OR ch > '9' THEN
            valid := FALSE;
        END_IF;
    END_FOR;

    FOR i := 1 TO TO_INT(seg2Len) DO
        ch := MID(seg2, 1, TO_INT(i));
        IF ch < '0' OR ch > '9' THEN
            valid := FALSE;
        END_IF;
    END_FOR;

    FOR i := 1 TO TO_INT(seg3Len) DO
        ch := MID(seg3, 1, TO_INT(i));
        IF ch < '0' OR ch > '9' THEN
            valid := FALSE;
        END_IF;
    END_FOR;

    FOR i := 1 TO TO_INT(seg4Len) DO
        ch := MID(seg4, 1, TO_INT(i));
        IF ch < '0' OR ch > '9' THEN
            valid := FALSE;
        END_IF;
    END_FOR;
END_IF;

IF valid THEN
    IF val1 <= 255 AND val2 <= 255 AND val3 <= 255 AND val4 <= 255 THEN
        result := (val1 * 16#1000000) OR (val2 * 16#10000) OR (val3 * 16#100) OR val4;
    END_IF;
END_IF;

ipValue := result;
END_FUNCTION_BLOCK

(* ---- public-medium-08.raw_candidate_01.st ---- *)
FUNCTION_BLOCK FB_ParseIPv4
VAR_INPUT
    ipText : STRING(254);
END_VAR
VAR_OUTPUT
    ipValue : UDINT;
END_VAR
VAR
    i : UINT;
    dot1 : UINT;
    dot2 : UINT;
    dot3 : UINT;
    len : UINT;
    seg1 : STRING(4);
    seg2 : STRING(4);
    seg3 : STRING(4);
    seg4 : STRING(4);
    seg1Len : UINT;
    seg2Len : UINT;
    seg3Len : UINT;
    seg4Len : UINT;
    val1 : UDINT;
    val2 : UDINT;
    val3 : UDINT;
    val4 : UDINT;
    result : UDINT;
    valid : BOOL;
    ch : CHAR;
END_VAR

result := 0;
valid := TRUE;

len := LEN(ipText);

IF len = 0 OR len > 254 THEN
    valid := FALSE;
END_IF

IF valid THEN
    dot1 := FIND(ipText, '.');
    IF dot1 <= 1 OR dot1 >= 254 THEN
        valid := FALSE;
    END_IF
END_IF

IF valid THEN
    dot2 := FIND(MID(ipText, 254 - dot1, dot1 + 1), '.');
    IF dot2 > 0 THEN
        dot2 := dot2 + dot1;
    END_IF;
END_IF;

IF valid THEN
    dot3 := 0;
    IF dot2 > 0 AND dot2 < 254 THEN
        dot3 := FIND(MID(ipText, 254 - dot2, dot2 + 1), '.');
        IF dot3 > 0 THEN
            dot3 := dot3 + dot2;
        END_IF;
    END_IF;
END_IF;

IF valid THEN
    IF dot1 = 0 OR dot2 = 0 OR dot3 = 0 THEN
        valid := FALSE;
    END_IF;
END_IF;

IF valid THEN
    seg1Len := dot1 - 1;
    seg2Len := dot2 - dot1 - 1;
    seg3Len := dot3 - dot2 - 1;
    seg4Len := len - dot3;

    IF seg1Len < 1 OR seg1Len > 3 OR seg2Len < 1 OR seg2Len > 3 OR
       seg3Len < 1 OR seg3Len > 3 OR seg4Len < 1 OR seg4Len > 3 THEN
        valid := FALSE;
    END_IF;
END_IF;

IF valid THEN
    seg1 := LEFT(ipText, seg1Len);
    seg2 := MID(ipText, seg2Len, dot1 + 1);
    seg3 := MID(ipText, seg3Len, dot2 + 1);
    seg4 := RIGHT(ipText, seg4Len);

    valid := (seg1Len = LEN(seg1)) AND (seg2Len = LEN(seg2)) AND
             (seg3Len = LEN(seg3)) AND (seg4Len = LEN(seg4));
END_IF;

IF valid THEN
    valid := FALSE;
    val1 := STRING_TO_UDINT(seg1);
    val2 := STRING_TO_UDINT(seg2);
    val3 := STRING_TO_UDINT(seg3);
    val4 := STRING_TO_UDINT(seg4);

    FOR i := 1 TO seg1Len DO
        ch := MID(seg1, 1, i);
        IF (ch < '0') OR (ch > '9') THEN
            valid := TRUE;
        END_IF;
    END_FOR;

    IF NOT valid THEN
        FOR i := 1 TO seg2Len DO
            ch := MID(seg2, 1, i);
            IF (ch < '0') OR (ch > '9') THEN
                valid := TRUE;
            END_IF;
        END_FOR;
    END_IF;

    IF NOT valid THEN
        FOR i := 1 TO seg3Len DO
            ch := MID(seg3, 1, i);
            IF (ch < '0') OR (ch > '9') THEN
                valid := TRUE;
            END_IF;
        END_FOR;
    END_IF;

    IF NOT valid THEN
        FOR i := 1 TO seg4Len DO
            ch := MID(seg4, 1, i);
            IF (ch < '0') OR (ch > '9') THEN
                valid := TRUE;
            END_IF;
        END_FOR;
    END_IF;

    IF valid THEN
        valid := FALSE;
    END_IF;
END_IF;

IF valid THEN
    IF val1 <= 255 AND val2 <= 255 AND val3 <= 255 AND val4 <= 255 THEN
        result := (val1 * 16#1000000) OR (val2 * 16#10000) OR (val3 * 16#100) OR val4;
    END_IF;
END_IF;

ipValue := result;
END_FUNCTION_BLOCK

(* ---- public-medium-08.raw_candidate_02.st ---- *)
FUNCTION_BLOCK FB_ParseIPv4
VAR_INPUT
    ipText : STRING(254);
END_VAR
VAR_OUTPUT
    ipValue : UDINT;
END_VAR
VAR
    i : UINT;
    dot1 : UINT;
    dot2 : UINT;
    dot3 : UINT;
    len : UINT;
    seg1 : STRING(4);
    seg2 : STRING(4);
    seg3 : STRING(4);
    seg4 : STRING(4);
    seg1Len : UINT;
    seg2Len : UINT;
    seg3Len : UINT;
    seg4Len : UINT;
    val1 : UDINT;
    val2 : UDINT;
    val3 : UDINT;
    val4 : UDINT;
    result : UDINT;
    valid : BOOL;
    ch : STRING(1);
END_VAR

result := 0;
valid := TRUE;

len := TO_UINT(LEN(ipText));

IF len = 0 OR len > 15 THEN
    valid := FALSE;
END_IF;

IF valid THEN
    dot1 := TO_UINT(FIND(ipText, '.'));
    IF dot1 <= 1 OR dot1 >= 254 THEN
        valid := FALSE;
    END_IF;
END_IF;

IF valid THEN
    dot2 := TO_UINT(FIND(MID(ipText, TO_INT(len - dot1), TO_INT(dot1 + 1)), '.'));
    IF dot2 > 0 THEN
        dot2 := dot2 + dot1;
    END_IF;
END_IF;

IF valid THEN
    dot3 := 0;
    IF dot2 > 0 AND dot2 < 254 THEN
        dot3 := TO_UINT(FIND(MID(ipText, TO_INT(len - dot2), TO_INT(dot2 + 1)), '.'));
        IF dot3 > 0 THEN
            dot3 := dot3 + dot2;
        END_IF;
    END_IF;
END_IF;

IF valid THEN
    IF dot1 = 0 OR dot2 = 0 OR dot3 = 0 THEN
        valid := FALSE;
    END_IF;
END_IF;

IF valid THEN
    seg1Len := dot1 - 1;
    seg2Len := dot2 - dot1 - 1;
    seg3Len := dot3 - dot2 - 1;
    seg4Len := len - dot3;

    IF seg1Len < 1 OR seg1Len > 3 OR seg2Len < 1 OR seg2Len > 3 OR seg3Len < 1 OR seg3Len > 3 OR seg4Len < 1 OR seg4Len > 3 THEN
        valid := FALSE;
    END_IF;
END_IF;

IF valid THEN
    seg1 := LEFT(ipText, TO_INT(seg1Len));
    seg2 := MID(ipText, TO_INT(seg2Len), TO_INT(dot1 + 1));
    seg3 := MID(ipText, TO_INT(seg3Len), TO_INT(dot2 + 1));
    seg4 := RIGHT(ipText, TO_INT(seg4Len));

    IF TO_UINT(LEN(seg1)) <> seg1Len OR TO_UINT(LEN(seg2)) <> seg2Len OR
       TO_UINT(LEN(seg3)) <> seg3Len OR TO_UINT(LEN(seg4)) <> seg4Len THEN
        valid := FALSE;
    END_IF;
END_IF;

IF valid THEN
    val1 := STRING_TO_UDINT(seg1);
    val2 := STRING_TO_UDINT(seg2);
    val3 := STRING_TO_UDINT(seg3);
    val4 := STRING_TO_UDINT(seg4);

    FOR i := 1 TO TO_INT(seg1Len) DO
        ch := MID(seg1, 1, TO_INT(i));
        IF ch < '0' OR ch > '9' THEN
            valid := FALSE;
        END_IF;
    END_FOR;

    FOR i := 1 TO TO_INT(seg2Len) DO
        ch := MID(seg2, 1, TO_INT(i));
        IF ch < '0' OR ch > '9' THEN
            valid := FALSE;
        END_IF;
    END_FOR;

    FOR i := 1 TO TO_INT(seg3Len) DO
        ch := MID(seg3, 1, TO_INT(i));
        IF ch < '0' OR ch > '9' THEN
            valid := FALSE;
        END_IF;
    END_FOR;

    FOR i := 1 TO TO_INT(seg4Len) DO
        ch := MID(seg4, 1, TO_INT(i));
        IF ch < '0' OR ch > '9' THEN
            valid := FALSE;
        END_IF;
    END_FOR;
END_IF;

IF valid THEN
    IF val1 <= 255 AND val2 <= 255 AND val3 <= 255 AND val4 <= 255 THEN
        result := (val1 * 16#1000000) OR (val2 * 16#10000) OR (val3 * 16#100) OR val4;
    END_IF;
END_IF;

ipValue := result;
END_FUNCTION_BLOCK

(* ---- self-easy-01.candidate_01.st ---- *)
FUNCTION_BLOCK FB
VAR
    lastAvgOut : REAL := 0.0;
END_VAR
VAR_OUTPUT
    avgOut : REAL := 0.0;
END_VAR
VAR_INPUT
    enable      : BOOL;
    values      : ARRAY[1..8] OF INT;
    count       : INT;
    avgEnable   : BOOL;
END_VAR
VAR
    sum   : DINT;
    i     : INT;
    n     : INT;
END_VAR

// [S2] enable = FALSE: keep previous
// [S5] avgEnable = FALSE: keep previous
// [S1] count <= 0: keep previous, avoid div-by-zero
// Guard: only compute when all conditions satisfied
IF enable AND avgEnable AND (count > 0) THEN
    // [S6] clamp count to array bounds [1..8]
    IF count > 8 THEN
        n := 8;
    ELSE
        n := count;
    END_IF;

    // Wide-type sum to prevent INT overflow
    sum := 0;
    FOR i := 1 TO n DO
        sum := sum + values[i];
    END_FOR;

    // [S4][S6] REAL division preserves fractional precision
    avgOut := DINT_TO_REAL(sum) / DINT_TO_REAL(n);
    lastAvgOut := avgOut;
ELSE
    avgOut := lastAvgOut;
END_IF;
END_FUNCTION_BLOCK

(* ---- self-easy-01.raw_candidate_01.st ---- *)
FUNCTION_BLOCK FB
VAR
    lastAvgOut : REAL := 0.0;
END_VAR
VAR_OUTPUT
    avgOut : REAL := 0.0;
END_VAR
VAR_INPUT
    enable      : BOOL;
    values      : ARRAY[1..8] OF INT;
    count       : INT;
    avgEnable   : BOOL;
END_VAR
VAR
    sum   : DINT;
    i     : INT;
    n     : INT;
END_VAR

// [S2] enable = FALSE: keep previous
// [S5] avgEnable = FALSE: keep previous
// [S1] count <= 0: keep previous, avoid div-by-zero
// Guard: only compute when all conditions satisfied
IF enable AND avgEnable AND (count > 0) THEN
    // [S6] clamp count to array bounds [1..8]
    IF count > 8 THEN
        n := 8;
    ELSE
        n := count;
    END_IF;

    // Wide-type sum to prevent INT overflow
    sum := 0;
    FOR i := 1 TO n DO
        sum := sum + values[i];
    END_FOR;

    // [S4][S6] REAL division preserves fractional precision
    avgOut := DINT_TO_REAL(sum) / DINT_TO_REAL(n);
    lastAvgOut := avgOut;
ELSE
    avgOut := lastAvgOut;
END_IF;
END_FUNCTION_BLOCK

(* ---- self-easy-02.candidate_01.st ---- *)
FUNCTION_BLOCK FB
VAR_INPUT
    tankLevel   : REAL;
    outletFlow  : REAL;
    inletPermit : BOOL;
    resetBtn    : BOOL;
END_VAR
VAR_OUTPUT
    pumpRun         : BOOL;
    alarmHigh       : BOOL;
    alarmLow        : BOOL;
    outletValveOpen : BOOL;
END_VAR
VAR
    prevResetBtn : BOOL := FALSE;
    latchHigh    : BOOL := FALSE;
    latchLow     : BOOL := FALSE;
END_VAR
VAR_TEMP
    risingReset : BOOL;
END_VAR

// Detect rising edge of reset button
risingReset := resetBtn AND NOT prevResetBtn;

// High level alarm: >= 85.0 sets immediately; falling below 85.0 clears only on rising reset
IF tankLevel >= 85.0 THEN
    latchHigh := TRUE;
ELSIF risingReset THEN
    latchHigh := FALSE;
END_IF;

// Low level alarm: <= 15.0 sets immediately; rising above 15.0 clears only on rising reset
IF tankLevel <= 15.0 THEN
    latchLow := TRUE;
ELSIF risingReset THEN
    latchLow := FALSE;
END_IF;

// Update latched states to outputs
alarmHigh := latchHigh;
alarmLow  := latchLow;

// Pump runs only when inlet permit is true AND both alarms are cleared
pumpRun := inletPermit AND (NOT alarmHigh) AND (NOT alarmLow);

// Outlet valve: open when low alarm is NOT latched
outletValveOpen := NOT alarmLow;

// Store button state for next scan edge detection
prevResetBtn := resetBtn;
END_FUNCTION_BLOCK

(* ---- self-easy-02.raw_candidate_01.st ---- *)
FUNCTION_BLOCK FB
VAR_INPUT
    tankLevel   : REAL;
    outletFlow  : REAL;
    inletPermit : BOOL;
    resetBtn    : BOOL;
END_VAR
VAR_OUTPUT
    pumpRun         : BOOL;
    alarmHigh       : BOOL;
    alarmLow        : BOOL;
    outletValveOpen : BOOL;
END_VAR
VAR
    prevResetBtn : BOOL := FALSE;
    latchHigh    : BOOL := FALSE;
    latchLow     : BOOL := FALSE;
END_VAR
VAR_TEMP
    risingReset : BOOL;
END_VAR

// Detect rising edge of reset button
risingReset := resetBtn AND NOT prevResetBtn;

// High level alarm: >= 85.0 sets immediately; falling below 85.0 clears only on rising reset
IF tankLevel >= 85.0 THEN
    latchHigh := TRUE;
ELSIF risingReset THEN
    latchHigh := FALSE;
END_IF;

// Low level alarm: <= 15.0 sets immediately; rising above 15.0 clears only on rising reset
IF tankLevel <= 15.0 THEN
    latchLow := TRUE;
ELSIF risingReset THEN
    latchLow := FALSE;
END_IF;

// Update latched states to outputs
alarmHigh := latchHigh;
alarmLow  := latchLow;

// Pump runs only when inlet permit is true AND both alarms are cleared
pumpRun := inletPermit AND (NOT alarmHigh) AND (NOT alarmLow);

// Outlet valve: open when low alarm is NOT latched
outletValveOpen := NOT alarmLow;

// Store button state for next scan edge detection
prevResetBtn := resetBtn;
END_FUNCTION_BLOCK

(* ---- self-hard-01.candidate_01.st ---- *)
FUNCTION_BLOCK FB
VAR_INPUT
    flowLow  : BOOL;
    ackBtn   : BOOL;
    sensorOK : BOOL;
END_VAR
VAR_OUTPUT
    alarmActive : BOOL;
    alarmAcked  : BOOL;
    highHigh    : BOOL;
END_VAR
VAR
    state        : UINT := 0;  // 0=IDLE, 1=UNACKED, 2=PENDING_CLEAR
    prevAckBtn   : BOOL := FALSE;
    prevFlowLow  : BOOL := FALSE;
    prevAlarmActive  : BOOL := FALSE;
    prevAlarmAcked   : BOOL := FALSE;
    risingEdge   : BOOL;   // rising edge of ackBtn
    risingEdge2  : BOOL;   // rising edge of flowLow
END_VAR

    // Edge detection
    risingEdge  := ackBtn AND NOT prevAckBtn;
    risingEdge2 := flowLow AND NOT prevFlowLow;

    // Update previous-cycle outputs for formal-property checks
    prevAlarmActive := alarmActive;
    prevAlarmAcked  := alarmAcked;

    // High-priority alarm: sensor failure
    highHigh := NOT sensorOK;

    // State machine
    CASE state OF
        0:  // IDLE
            alarmActive := FALSE;
            alarmAcked  := FALSE;
            IF risingEdge2 THEN
                state       := 1;
                alarmActive := TRUE;
                alarmAcked  := FALSE;
            ELSIF risingEdge AND flowLow THEN
                state       := 1;
                alarmActive := TRUE;
                alarmAcked  := FALSE;
            END_IF;

        1:  // UNACKED
            alarmActive := TRUE;
            alarmAcked  := FALSE;
            IF risingEdge2 THEN
                state := 1;  // re-triggered; remain UNACKED
            ELSIF risingEdge THEN
                state := 0;  // acked while condition still present
            ELSIF NOT flowLow THEN
                state       := 2;
                alarmAcked  := TRUE;  // condition gone, waiting for ack
            END_IF;

        2:  // PENDING_CLEAR
            alarmActive := TRUE;
            alarmAcked  := TRUE;
            IF risingEdge2 THEN
                state       := 1;
                alarmAcked  := FALSE;  // condition reappeared before ack
            ELSIF risingEdge THEN
                state       := 0;      // acked; condition already gone
                alarmActive := FALSE;
                alarmAcked  := FALSE;
            END_IF;
    END_CASE;

    // Shift register for next cycle edge detection
    prevAckBtn  := ackBtn;
    prevFlowLow := flowLow;
END_FUNCTION_BLOCK

(* ---- self-hard-01.candidate_02.st ---- *)
FUNCTION_BLOCK FB
VAR_INPUT
    flowLow  : BOOL;
    ackBtn   : BOOL;
    sensorOK : BOOL;
END_VAR
VAR_OUTPUT
    alarmActive : BOOL;
    alarmAcked  : BOOL;
    highHigh    : BOOL;
END_VAR
VAR
    prevAckBtn  : BOOL := FALSE;
    prevFlowLow : BOOL := FALSE;
    risingAck   : BOOL;
    risingFlow  : BOOL;
END_VAR

    // Rising edge detection
    risingAck  := ackBtn AND NOT prevAckBtn;
    risingFlow := flowLow AND NOT prevFlowLow;

    // High-priority: sensor failure
    highHigh := NOT sensorOK;

    // Main alarm logic
    IF risingFlow THEN
        // Condition reappeared → unacknowledged active alarm
        alarmActive := TRUE;
        alarmAcked  := FALSE;
    ELSIF risingAck THEN
        // Acknowledge button pressed
        IF flowLow THEN
            // Condition still present: acknowledge only
            alarmActive := TRUE;
            alarmAcked  := TRUE;
        ELSE
            // Condition already gone: clear alarm
            alarmActive := FALSE;
            alarmAcked  := FALSE;
        END_IF;
    ELSIF alarmActive AND NOT alarmAcked AND NOT flowLow THEN
        // Condition disappeared before acknowledgment → pending clear
        alarmActive := TRUE;
        alarmAcked  := TRUE;
    END_IF;

    prevAckBtn  := ackBtn;
    prevFlowLow := flowLow;
END_FUNCTION_BLOCK

(* ---- self-hard-01.raw_candidate_01.st ---- *)
FUNCTION_BLOCK FB
VAR_INPUT
    flowLow  : BOOL;
    ackBtn   : BOOL;
    sensorOK : BOOL;
END_VAR
VAR_OUTPUT
    alarmActive : BOOL;
    alarmAcked  : BOOL;
    highHigh    : BOOL;
END_VAR
VAR
    state        : UINT := 0;  // 0=IDLE, 1=UNACKED, 2=PENDING_CLEAR
    prevAckBtn   : BOOL := FALSE;
    prevFlowLow  : BOOL := FALSE;
    prevAlarmActive  : BOOL := FALSE;
    prevAlarmAcked   : BOOL := FALSE;
    risingEdge   : BOOL;   // rising edge of ackBtn
    risingEdge2  : BOOL;   // rising edge of flowLow
END_VAR

    // Edge detection
    risingEdge  := ackBtn AND NOT prevAckBtn;
    risingEdge2 := flowLow AND NOT prevFlowLow;

    // Update previous-cycle outputs for formal-property checks
    prevAlarmActive := alarmActive;
    prevAlarmAcked  := alarmAcked;

    // High-priority alarm: sensor failure
    highHigh := NOT sensorOK;

    // State machine
    CASE state OF
        0:  // IDLE
            alarmActive := FALSE;
            alarmAcked  := FALSE;
            IF risingEdge2 THEN
                state       := 1;
                alarmActive := TRUE;
                alarmAcked  := FALSE;
            ELSIF risingEdge AND flowLow THEN
                state       := 1;
                alarmActive := TRUE;
                alarmAcked  := FALSE;
            END_IF;

        1:  // UNACKED
            alarmActive := TRUE;
            alarmAcked  := FALSE;
            IF risingEdge2 THEN
                state := 1;  // re-triggered; remain UNACKED
            ELSIF risingEdge THEN
                state := 0;  // acked while condition still present
            ELSIF NOT flowLow THEN
                state       := 2;
                alarmAcked  := TRUE;  // condition gone, waiting for ack
            END_IF;

        2:  // PENDING_CLEAR
            alarmActive := TRUE;
            alarmAcked  := TRUE;
            IF risingEdge2 THEN
                state       := 1;
                alarmAcked  := FALSE;  // condition reappeared before ack
            ELSIF risingEdge THEN
                state       := 0;      // acked; condition already gone
                alarmActive := FALSE;
                alarmAcked  := FALSE;
            END_IF;
    END_CASE;

    // Shift register for next cycle edge detection
    prevAckBtn  := ackBtn;
    prevFlowLow := flowLow;
END_FUNCTION_BLOCK

(* ---- self-hard-01.raw_candidate_02.st ---- *)
FUNCTION_BLOCK FB
VAR_INPUT
    flowLow  : BOOL;
    ackBtn   : BOOL;
    sensorOK : BOOL;
END_VAR
VAR_OUTPUT
    alarmActive : BOOL;
    alarmAcked  : BOOL;
    highHigh    : BOOL;
END_VAR
VAR
    prevAckBtn  : BOOL := FALSE;
    prevFlowLow : BOOL := FALSE;
    risingAck   : BOOL;
    risingFlow  : BOOL;
END_VAR

    // Rising edge detection
    risingAck  := ackBtn AND NOT prevAckBtn;
    risingFlow := flowLow AND NOT prevFlowLow;

    // High-priority: sensor failure
    highHigh := NOT sensorOK;

    // Main alarm logic
    IF risingFlow THEN
        // Condition reappeared → unacknowledged active alarm
        alarmActive := TRUE;
        alarmAcked  := FALSE;
    ELSIF risingAck THEN
        // Acknowledge button pressed
        IF flowLow THEN
            // Condition still present: acknowledge only
            alarmActive := TRUE;
            alarmAcked  := TRUE;
        ELSE
            // Condition already gone: clear alarm
            alarmActive := FALSE;
            alarmAcked  := FALSE;
        END_IF;
    ELSIF alarmActive AND NOT alarmAcked AND NOT flowLow THEN
        // Condition disappeared before acknowledgment → pending clear
        alarmActive := TRUE;
        alarmAcked  := TRUE;
    END_IF;

    prevAckBtn  := ackBtn;
    prevFlowLow := flowLow;
END_FUNCTION_BLOCK

(* ---- self-hard-02.candidate_01.st ---- *)
FUNCTION_BLOCK FB
VAR_INPUT
    startBtn   : BOOL;
    abortBtn   : BOOL;
    setpoint   : REAL;
    pv         : REAL;
    maxDuration: INT;
END_VAR
VAR_OUTPUT
    elapsed : INT := 0;
    phase   : INT := 0;
    timeout : BOOL := FALSE;
END_VAR
VAR
    prev_startBtn : BOOL := FALSE;
    prev_phase    : INT  := 0;
    risingEdge    : BOOL;
END_VAR

    // Detect rising edge of startBtn before any state changes this scan
    risingEdge := startBtn AND NOT prev_startBtn;

    // Priority 1: abort
    IF abortBtn THEN
        phase   := 9;
        // elapsed and timeout stay frozen (no assignment)

    // Priority 2: new rising edge (only if not aborted this scan)
    ELSIF risingEdge THEN
        elapsed := 0;
        timeout := FALSE;
        phase   := 1;

    // Priority 3: running phases — count and evaluate transition
    ELSIF (prev_phase = 1) OR (prev_phase = 2) THEN
        elapsed := elapsed + 1;

        // Check timeout before setting phase
        IF elapsed >= maxDuration THEN
            timeout := TRUE;
            phase   := 3;
        ELSE
            // Phase transition based on temperature
            IF (prev_phase = 2) OR (pv >= setpoint) THEN
                phase := 2;
            ELSE
                phase := 1;
            END_IF;
        END_IF;

    // Frozen states (phase 0, 3, 9) — no changes to elapsed/phase/timeout
    ELSE
        // phase, elapsed, timeout retain their values
    END_IF;

    // Update previous-cycle snapshot for next scan
    prev_startBtn := startBtn;
    prev_phase    := phase;
END_FUNCTION_BLOCK

(* ---- self-hard-02.candidate_02.st ---- *)
FUNCTION_BLOCK FB
VAR_INPUT
    startBtn   : BOOL;
    abortBtn   : BOOL;
    setpoint   : REAL;
    pv         : REAL;
    maxDuration: INT;
END_VAR
VAR_OUTPUT
    elapsed  : INT  := 0;
    phase    : INT  := 0;
    timeout  : BOOL := FALSE;
END_VAR
VAR
    prev_startBtn : BOOL := FALSE;
    prev_phase    : INT  := 0;
    risingEdge    : BOOL;
END_VAR

    risingEdge := startBtn AND NOT prev_startBtn;

    IF abortBtn THEN
        phase := 9;
        elapsed := elapsed;
        timeout := timeout;

    ELSIF risingEdge THEN
        elapsed := 0;
        timeout := FALSE;
        phase   := 1;

    ELSIF (prev_phase = 1) OR (prev_phase = 2) THEN
        elapsed := elapsed + 1;

        IF elapsed >= maxDuration THEN
            timeout := TRUE;
            phase   := 3;
        ELSE
            IF (prev_phase = 2) OR (pv >= setpoint) THEN
                phase := 2;
            ELSE
                phase := 1;
            END_IF;
        END_IF;

    ELSE
        NULL;
    END_IF;

    prev_startBtn := startBtn;
    prev_phase    := phase;
END_FUNCTION_BLOCK
